(* Logix 5000 project; controller TFF vendor 1 type 14 code 107 rev 34.11; software revision 34.03; part 20 of 36 *)
(* tags used below, declared in another part *)
   Address : DINT;   // Temp Address
   Config : Configuration;   // Index Array used in configuration routines
   Index : DINT;   // Index
   NewSystem : DINT;
   AI101 : ALIAS FOR AnalogPoint[10];   // Filtrate Conductivity
   AI101_SIG : ALIAS FOR DigitalPoint[90];
   AI102 : ALIAS FOR AnalogPoint[11];   // Filtrate UV
   AI102_SIG : ALIAS FOR DigitalPoint[91];
   AI103 : ALIAS FOR AnalogPoint[12];   // Filtrate UV
   AI103_SIG : ALIAS FOR DigitalPoint[92];
   AI104 : ALIAS FOR AnalogPoint[9];   // Filtrate pH
   AI104_SIG : ALIAS FOR DigitalPoint[105];
   AlarmAnalog : AlarmAnalog[50];   // Analog Alarm Array
   AlarmControl : AlarmControl;   // Alarm Control
   AlarmDeviation : AlarmDeviation[20];   // Control Loop Deviation Alarm Array
   AnalogOutput : AnalogOutput[25];   // Analog Output Array
   AnalogPoint : AnalogInput[50];   // Analog Input Array
   Concentration : Concentration;
   ControlLoop : ControlLoop[20];   // Control Loop Array
   ControlLoop_FeedBagLevel : ALIAS FOR ControlLoop[2];   // Feed Bag Level Control Loop
   Diafiltration : Diafiltration;
   DigitalOutput : BOOL[256];   // Digital Output Array these bits are sent to output cards.
   DigitalPoint : DigitalPoint[150];   // Digital Point Array
   DP : ALIAS FOR AnalogPoint[40];   // Differential Pressure
   Drive : Drive[11];   // Drives Array
   ES001 : ALIAS FOR DigitalPoint[3];   // Emergency Stop
   FI001 : ALIAS FOR AnalogPoint[42];   // Feed Flow
   FI003 : ALIAS FOR AnalogPoint[17];
   FI003_SIG : ALIAS FOR DigitalPoint[106];
   FI003Alarm : ALIAS FOR AlarmAnalog[17];
   FI101 : ALIAS FOR AnalogPoint[2];   // Filtrate Flow
   FI101_SIG : ALIAS FOR DigitalPoint[93];
   FI101Alarm : ALIAS FOR AlarmAnalog[2];   // Filtrate Flow Alarm
   FI401 : ALIAS FOR AnalogPoint[43];   // Transfer Pump Flow
   LI001 : ALIAS FOR AnalogPoint[44];   // Feed Bag Volume
   LI001Alarm : ALIAS FOR AlarmAnalog[44];   // Feed Bag Volume Alarm
   MIX001 : ALIAS FOR AnalogPoint[14];   // Mixer Speed
   MIX001_SIG : ALIAS FOR DigitalPoint[104];
   Mixer : Mixer;   // Mixer config. structure
   NWP : ALIAS FOR AnalogPoint[45];   // Normalized Water Permeability
   Options : Options;   // Options List
   PCV001 : ALIAS FOR AnalogPoint[3];   // Retentate Pressure Control Valve Position
   PCV001_Control : PCV_Control;   // PCV001 Control UDT
   PCV001_SIG : ALIAS FOR DigitalPoint[102];
   PCV101 : ALIAS FOR AnalogPoint[4];   // Filtrate Pressure Control Valve Position
   PCV101_Control : PCV_Control;   // PCV101 Control UDT
   PCV101_SIG : ALIAS FOR DigitalPoint[103];
   PERM : ALIAS FOR AnalogPoint[46];   // Membrane Permeability
   PI001 : ALIAS FOR AnalogPoint[5];   // Feed Pressure
   PI001_SIG : ALIAS FOR DigitalPoint[97];
   PI002 : ALIAS FOR AnalogPoint[6];   // Retentate Pressure
   PI002_SIG : ALIAS FOR DigitalPoint[98];
   PI101 : ALIAS FOR AnalogPoint[7];   // Filtrate Pressure
   PI101_SIG : ALIAS FOR DigitalPoint[99];
   PI401 : ALIAS FOR AnalogPoint[8];   // Transfer Pump Pressure
   PI401_SIG : ALIAS FOR DigitalPoint[100];
   PSH001 : ALIAS FOR DigitalPoint[4];   // Feed Pump High Pressure
   PSH401 : ALIAS FOR DigitalPoint[5];   // Transfer Pump High Pressure
   PSL602 : ALIAS FOR DigitalPoint[0];   // Valves Air Defect
   PSL603 : ALIAS FOR DigitalPoint[10];   // Manifold Valves Air Defect
   SIC001 : ALIAS FOR Drive[1];   // Feed Pump
   SIC001DF : ALIAS FOR DigitalPoint[8];   // Feed Pump Defect
   SIC002 : ALIAS FOR Drive[2];   // Transfer Pump
   SIC002DF : ALIAS FOR DigitalPoint[9];   // Transfer Pump Defect
   SIC003 : ALIAS FOR Drive[3];   // Mixer
   SIC003DF : ALIAS FOR DigitalPoint[14];   // Mixer Defect
   SRL001 : ALIAS FOR DigitalPoint[15];   // Tank Skid Remote / Standalone
   Tank : TankManagement;   // Tank Management
   ThisSystem : SystemType;
   TI001 : ALIAS FOR AnalogPoint[13];   // Feed Bag Temperature
   TI001_SIG : ALIAS FOR DigitalPoint[101];
   TMP : ALIAS FOR AnalogPoint[41];   // Trans-membrane Pressure
   Totalizer : Totalizers[20];   // Totalizers Array
   UserCr1 : ALIAS FOR DigitalPoint[65];   // User Critical Alarm 1
   UserCr2 : ALIAS FOR DigitalPoint[67];   // User Critical Alarm 2
   UserNCr1 : ALIAS FOR DigitalPoint[64];   // User Non Critical Alarm 1
   UserNCr2 : ALIAS FOR DigitalPoint[66];   // User Non Critical Alarm 2
   Valve : Valve[100];   // Valve Array
   WI001 : ALIAS FOR AnalogPoint[15];   // Feed Bag Weight
   WI001_SIG : ALIAS FOR DigitalPoint[94];
   WI001Alarm : ALIAS FOR AlarmAnalog[15];   // Feed Bag Weight Alarm
   WI101 : ALIAS FOR AnalogPoint[0];   // Filtrate Weight
   WI101_SIG : ALIAS FOR DigitalPoint[95];
   WI101Alarm : ALIAS FOR AlarmAnalog[0];   // Filtrate Weight Alarm
   WI102 : ALIAS FOR AnalogPoint[1];   // Customer Filtrate Weight
   WI102_SIG : ALIAS FOR DigitalPoint[96];
   WI102Alarm : ALIAS FOR AlarmAnalog[1];   // Customer Filtrate Weight Alarm
   XC102_3DF : ALIAS FOR DigitalPoint[13];   // C8000 Defect
   XS001 : ALIAS FOR DigitalPoint[1];   // Door Closed
   XS002 : ALIAS FOR DigitalPoint[6];   // Clamshell Locking 1 Closed
   XS003 : ALIAS FOR DigitalPoint[7];   // Clamshell Locking 2 Closed
   XS006 : ALIAS FOR DigitalPoint[2];   // Door to Frame Locking Closed
   XS011 : ALIAS FOR DigitalPoint[11];   // Pump P001 Type
   XS012 : ALIAS FOR DigitalPoint[12];   // Pump P002 Type
   YA01 : ALIAS FOR DigitalPoint[50];   // PC to PLC communication failure
   YA02 : ALIAS FOR DigitalPoint[51];   // CCP Runtime communication failure
   YA03 : ALIAS FOR DigitalPoint[52];   // Historical Data collection failure
   YA04 : ALIAS FOR DigitalPoint[53];   // Hard Drive Overload
   YA05 : ALIAS FOR DigitalPoint[54];   // Database Overload
   YA06 : ALIAS FOR DigitalPoint[55];   // Node 0 communication failure - Smart
   YA07 : ALIAS FOR DigitalPoint[56];   // Node 0 internal defect - Smart
   YA08 : ALIAS FOR DigitalPoint[57];   // Node 1 communication failure - Clamshell
   YA09 : ALIAS FOR DigitalPoint[58];   // Node 1 internal defect - Clamshell
   YA10 : ALIAS FOR DigitalPoint[59];   // PLC Program Major Fault
   YA11 : ALIAS FOR DigitalPoint[60];   // Database Corrupted
   YA12 : ALIAS FOR DigitalPoint[61];   // Unauthorized accesses
   YA13 : ALIAS FOR DigitalPoint[62];   // Tank Size Mismatch
   YA14 : ALIAS FOR DigitalPoint[63];   // SQL Server Write Failure
   YA15 : ALIAS FOR DigitalPoint[69];   // Node 3 Communication Failure - Pump
   YA16 : ALIAS FOR DigitalPoint[70];   // Node 3 Internal Defect - Pump
   YA17 : ALIAS FOR DigitalPoint[71];   // Node 4 Communication Failure - Instrum
   YA18 : ALIAS FOR DigitalPoint[72];   // Node 4 Internal Defect - Instrum
   YA19 : ALIAS FOR DigitalPoint[73];   // Node 5 Communication Failure - Tank
   YA20 : ALIAS FOR DigitalPoint[74];   // Node 5 Internal Defect - Tank
   YA21 : ALIAS FOR DigitalPoint[75];   // Node 6 IND331 Communication Failure
   YA22 : ALIAS FOR DigitalPoint[76];   // Node 7 IND131 Communication Failure
   YA41 : ALIAS FOR DigitalPoint[77];   // YA41 Operating Time Exceeded
   ZSDF : ALIAS FOR DigitalPoint[68];   // ZSDF Clamshell Locking Defect
(* Process, continued *)

ROUTINE Alarm_Init_Config   (* structured text *)
   (* =======================================================================
   	Alarm_Init_SP : initialized  parameter to default values
   
   	List of treatments
   		- Analog alarms set point with scale Min and Max
   		- Deviation alarms
   		- Digital alarmss
   		- Valves alarms
   	-----------------------------------------------------------------------------------------------------------------------------------------------------
   	History
   		2020-Sep-28 - Merck - Q.Spindler - Initial version for Candidate Release 3.00.00.01.a
   		2021-May-31 - DAVIDSON- Ch. ARBOGAST - Modifications for Candidate Release 3.01.00.00.a
   		On Analog Set point, add lines for set WI001 & LI001, HI & HIHI values according to actual tank size
   		On Analog Set point, add lines for set WI101 & WI102 & FI003 & FI101, HI & HIHI values according to actual system type
   		On Discrete Alarms: modify YA03.DelayTimerSP := 80
   		On Discrete Alarms: for all “_SIG” alarms, modify: Priority := 0 , DelayTimerSP := 10
   		On Discrete Alarms add line with WI001_SIG settings
   		On Discrete Alarms, last line FI003 settings: replace AI104 by FI003 (2x)
   =============================================================================================================================*)
   
   (*Analog Set point to min/max scale, Enable alarm, timer to  2s
   ============================================================*)
   	FOR Index := 0 to 49 by 1 do
   		IF AnalogPoint[Index].EnableCfg THEN
   			AlarmAnalog[Index].Override := 0; // Enable
   			AlarmAnalog[Index].LOLO := AnalogPoint[Index].ScaledMin ;
   			AlarmAnalog[Index].LO := AnalogPoint[Index].ScaledMin ;
   			AlarmAnalog[Index].HI := AnalogPoint[Index].ScaledMax ;
   			AlarmAnalog[Index].HIHI := AnalogPoint[Index].ScaledMax ;
   			AlarmAnalog[Index].LOLOTimerSP := 2 ;
   			AlarmAnalog[Index].LOTimerSP := 2 ;
   			AlarmAnalog[Index].HITimerSP := 2 ;
   			AlarmAnalog[Index].HIHITimerSP := 2 ;
   		END_IF;
   	End_for ;
   	(* Tank 60(50L) *)
   	IF Tank.Config.TankSelected = 1 THEN
   		WI001Alarm.HIHI := 60 ;
   		WI001Alarm.HI := 60 ;
   		LI001Alarm.HIHI := 50 ;
   		LI001Alarm.HI := 50 ;
   	END_IF ;
   	(* Tank 120(100L) *)
   	IF Tank.Config.TankSelected = 2 THEN
   		WI001Alarm.HIHI := 120 ;
   		WI001Alarm.HI := 120 ;
   		LI001Alarm.HIHI := 100 ;
   		LI001Alarm.HI := 100 ;
   	END_IF ;
   	(* Tank 240(200L) *)
   	IF Tank.Config.TankSelected = 3 THEN
   		WI001Alarm.HIHI := 240 ;
   		WI001Alarm.HI := 240 ;
   		LI001Alarm.HIHI := 200 ;
   		LI001Alarm.HI := 200 ;
   	END_IF ;
   	(* TF2S *)
   	IF NewSystem = 123 THEN
   		WI101Alarm.HIHI := 600 ;
   		WI101Alarm.HI := 600 ;
   		WI102Alarm.HIHI := 1000 ;
   		WI102Alarm.HI := 1000 ;
   		FI003Alarm.HIHI := 15 ;
   		FI003Alarm.HI := 15 ;
   		FI101Alarm.HIHI := 15 ;
   		FI101Alarm.HI := 15 ;
   	END_IF ;
   	(* TF3S *)
   	IF NewSystem = 124 THEN
   		WI101Alarm.HIHI := 1500 ;
   		WI101Alarm.HI := 1500 ;
   		WI102Alarm.HIHI := 1500 ;
   		WI102Alarm.HI := 1500 ;
   		FI003Alarm.HIHI := 25 ;
   		FI003Alarm.HI := 25 ;
   		FI101Alarm.HIHI := 25 ;
   		FI101Alarm.HI := 25 ;
   	END_IF ;
   
   (*Deviation alarm HI 100% HIHI 100%, Disable alarm, timer to 2s
   ============================================================*)
   	FOR Index := 0 to 19 by 1 do
   		IF AlarmDeviation[Index].EnableCfg THEN
   			AlarmDeviation[Index].Override := 1; // Disable
   			AlarmDeviation[Index].HI := 100 ;
   			AlarmDeviation[Index].HIHI := 100 ;
   			AlarmDeviation[Index].HITimerSP := 2 ;
   			AlarmDeviation[Index].HIHITImerSP := 2 ;
   		END_IF;
   	End_for ;
   
   (* Discrete Alarms
   ============================================================*)
   	ES001.DelayTimerSP := 0;
   	PSH001.Override := 0; PSH001.Priority := 1; PSH001.DelayTimerSP := 0;
   	PSH401.Override := 0; PSH401.Priority := 1; PSH401.DelayTimerSP := 0;
   	PSL602.Override := 0; PSL602.Priority := 1; PSL602.DelayTimerSP := 2;
   	SIC001DF.Override := 0; SIC001DF.Priority := 1; SIC001DF.DelayTimerSP :=1;
   	SIC002DF.Override := 0; SIC002DF.Priority := 1; SIC002DF.DelayTimerSP :=1;
   	SIC003DF.Override := 0; SIC003DF.Priority := 1; SIC003DF.DelayTimerSP :=1;
   	XC102_3DF.Override := 0; XC102_3DF.Priority := 1; XC102_3DF.DelayTimerSP :=1;
   	ZSDF.Override := 0; ZSDF.Priority := 1; ZSDF.DelayTimerSP :=1;
   	XS001.Override := 0; XS001.Priority := 1; XS001.DelayTimerSP :=1;
   	PSL603.Override := 0; PSL603.Priority := 1; PSL603.DelayTimerSP :=1;
   
   	YA01.Override := 0; YA01.Priority := 0; YA01.DelayTimerSP := 60;
   	YA02.Override := 0; YA02.Priority := 0; YA02.DelayTimerSP := 60;
   	YA03.Override := 0; YA03.Priority := 0; YA03.DelayTimerSP := 80;
   	YA04.Override := 0; YA04.Priority := 0; YA04.DelayTimerSP := 60;
   	YA05.Override := 0; YA05.Priority := 0; YA05.DelayTimerSP := 60;
   	YA06.Override := 0; YA06.Priority := 1; YA06.DelayTimerSP := 5;
   	YA07.Override := 0; YA07.Priority := 0; YA07.DelayTimerSP := 2;
   	YA08.Override := 0; YA08.Priority := 1; YA08.DelayTimerSP := 5;
   	YA09.Override := 0; YA09.Priority := 0; YA09.DelayTimerSP := 2;
   	YA10.DelayTimerSP := 0;
   	YA11.Override := 1; YA11.Priority := 0; YA11.DelayTimerSP := 5;
   	YA12.Override := 0; YA12.Priority := 0; YA12.DelayTimerSP := 0;
   	YA13.Override := 0; YA13.Priority := 0; YA13.DelayTimerSP := 2;
   	YA14.Override := 0; YA14.Priority := 0; YA14.DelayTimerSP := 60;
   	YA15.Override := 0; YA15.Priority := 1; YA15.DelayTimerSP := 5;
   	YA16.Override := 0; YA16.Priority := 0; YA16.DelayTimerSP := 2;
   	YA17.Override := 0; YA17.Priority := 1; YA17.DelayTimerSP := 5;
   	YA18.Override := 0; YA18.Priority := 0; YA18.DelayTimerSP := 2;
   	YA19.Override := 0; YA19.Priority := 1; YA19.DelayTimerSP := 5;
   	YA20.Override := 0; YA20.Priority := 0; YA20.DelayTimerSP := 2;
   	YA21.Override := 0; YA21.Priority := 1; YA21.DelayTimerSP := 5;
   	YA22.Override := 0; YA22.Priority := 1; YA22.DelayTimerSP := 5;
   
   	AI101_SIG.Override := 0; AI101_SIG.Priority := 0; AI101_SIG.DelayTimerSP := 10;
   	AI102_SIG.Override := 0; AI102_SIG.Priority := 0; AI102_SIG.DelayTimerSP := 10;
   	AI103_SIG.Override := 0; AI103_SIG.Priority := 0; AI103_SIG.DelayTimerSP := 10;
   	FI101_SIG.Override := 0; FI101_SIG.Priority := 0; FI101_SIG.DelayTimerSP := 10;
   	WI001_SIG.Override := 0; WI001_SIG.Priority := 0; WI001_SIG.DelayTimerSP := 10;
   	WI101_SIG.Override := 0; WI101_SIG.Priority := 0; WI101_SIG.DelayTimerSP := 10;
   	WI102_SIG.Override := 0; WI102_SIG.Priority := 0; WI102_SIG.DelayTimerSP := 10;
   	PI001_SIG.Override := 0; PI001_SIG.Priority := 0; PI001_SIG.DelayTimerSP := 10;
   	PI002_SIG.Override := 0; PI002_SIG.Priority := 0; PI002_SIG.DelayTimerSP := 10;
   	PI101_SIG.Override := 0; PI101_SIG.Priority := 0; PI101_SIG.DelayTimerSP := 10;
   	PI401_SIG.Override := 0; PI401_SIG.Priority := 0; PI401_SIG.DelayTimerSP := 10;
   	TI001_SIG.Override := 0; TI001_SIG.Priority := 0; TI001_SIG.DelayTimerSP := 10;
   	PCV001_SIG.Override := 0; PCV001_SIG.Priority := 0; PCV001_SIG.DelayTimerSP := 10;
   	PCV101_SIG.Override := 0; PCV101_SIG.Priority := 0; PCV101_SIG.DelayTimerSP := 10;
   	MIX001_SIG.Override := 0; MIX001_SIG.Priority := 0; MIX001_SIG.DelayTimerSP := 10;
   	AI104_SIG.Override := 0; AI104_SIG.Priority := 0; AI104_SIG.DelayTimerSP := 10;
   	FI003_SIG.Override := 0; FI003_SIG.Priority := 0; FI003_SIG.DelayTimerSP := 10;
   
   	UserNCr1.Priority := 0; UserNCr1.DelayTimerSP := 0;
   	UserCr1.Priority := 1; UserCr1.DelayTimerSP := 0;
   	UserNCr2.Priority := 0; UserNCr2.DelayTimerSP := 0;
   	UserCr2.Priority := 1; UserCr2.DelayTimerSP := 0;
   
   // Reset Init command
   AlarmControl.InitAlarmConfig := 0;
END_ROUTINE

ROUTINE Concentration_Diafiltration   (* ladder *)
// Agitator Control Routine
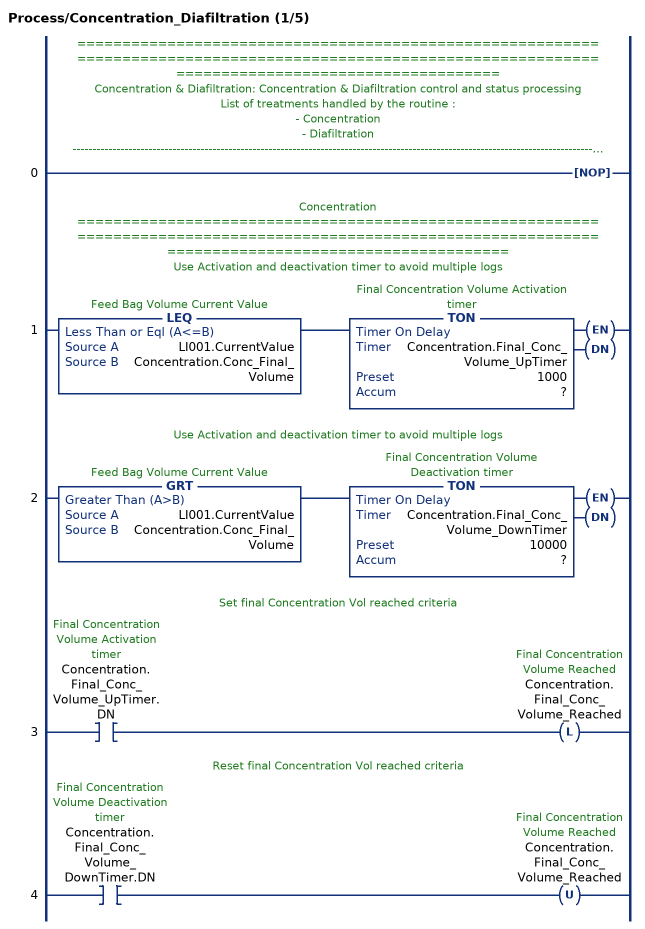
   // ========================================================================================================================================================
   //                                                                                                    Concentration & Diafiltration: Concentration & Diafiltration control and status processing
   //                                                     List of treatments handled by the routine :
   //                                                          - Concentration
   //                                                          - Diafiltration
   //                                                     -----------------------------------------------------------------------------------------------------------------------------------------------------
   //                                                     History
   //                                                          2019-AUG-13 - Actemium - B. Roch - Initial version for Candidate Release 3.00.00.00.a
   //                                                           2020-SEP-24 - Merck - Q. Spindler - Modifications for Candidate Release 3.00.00.01.a
   //                                        - Add Timer for activation and deactivation of Volume/Protein reached status to avoid unwanted logs
   // ========================================================================================================================================================
   0: NOP();
   // Concentration
   // ==========================================================================================================================================================
   // Use Activation and deactivation timer to avoid multiple logs
   1: LEQ(LI001.CurrentValue,Concentration.Conc_Final_Volume)TON(Concentration.Final_Conc_Volume_UpTimer,?,?);
   // Use Activation and deactivation timer to avoid multiple logs
   2: GRT(LI001.CurrentValue,Concentration.Conc_Final_Volume)TON(Concentration.Final_Conc_Volume_DownTimer,?,?);
   // Set final Concentration Vol reached criteria
   3: XIC(Concentration.Final_Conc_Volume_UpTimer.DN)OTL(Concentration.Final_Conc_Volume_Reached);
   // Reset final Concentration Vol reached criteria
   4: XIC(Concentration.Final_Conc_Volume_DownTimer.DN)OTU(Concentration.Final_Conc_Volume_Reached);
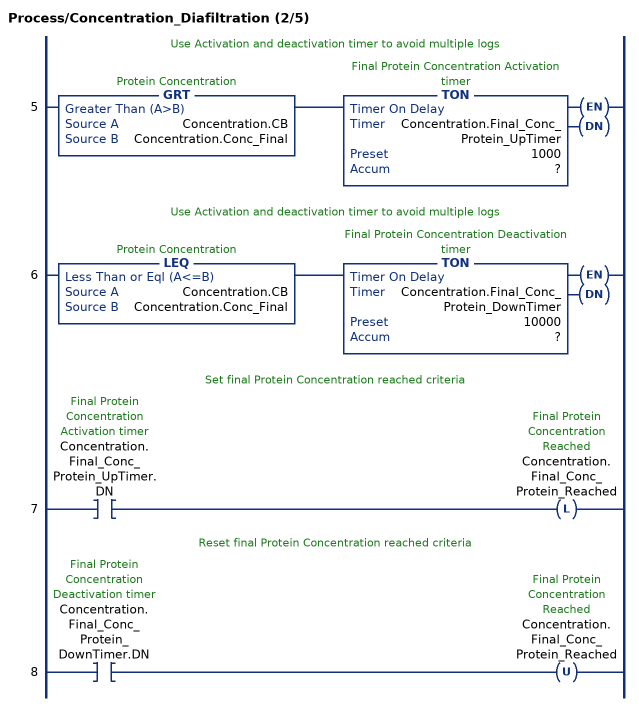
   // Use Activation and deactivation timer to avoid multiple logs
   5: GRT(Concentration.CB,Concentration.Conc_Final)TON(Concentration.Final_Conc_Protein_UpTimer,?,?);
   // Use Activation and deactivation timer to avoid multiple logs
   6: LEQ(Concentration.CB,Concentration.Conc_Final)TON(Concentration.Final_Conc_Protein_DownTimer,?,?);
   // Set final Protein Concentration reached criteria
   7: XIC(Concentration.Final_Conc_Protein_UpTimer.DN)OTL(Concentration.Final_Conc_Protein_Reached);
   // Reset final Protein Concentration reached criteria
   8: XIC(Concentration.Final_Conc_Protein_DownTimer.DN)OTU(Concentration.Final_Conc_Protein_Reached);
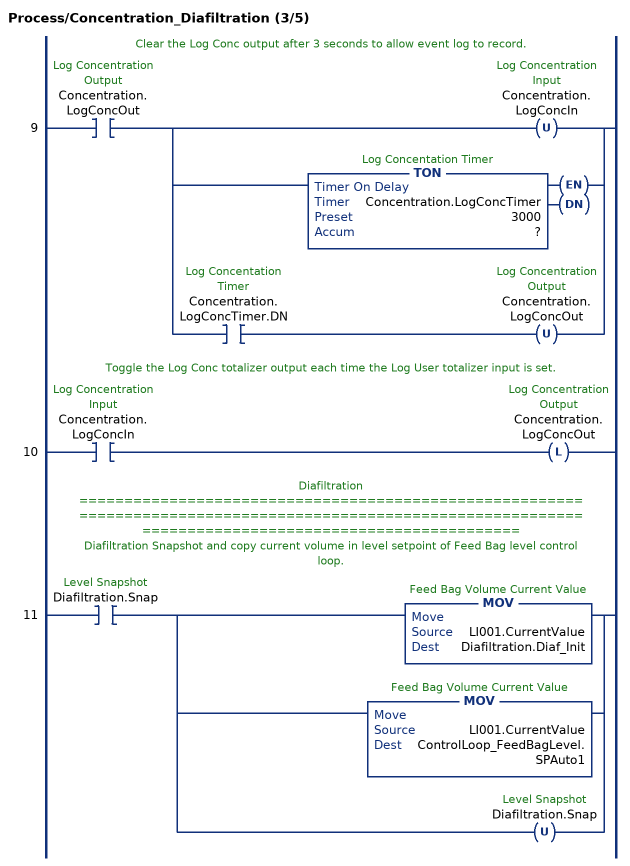
   // Clear the Log Conc output after 3 seconds to allow event log to record.
   9: XIC(Concentration.LogConcOut)[OTU(Concentration.LogConcIn) ,TON(Concentration.LogConcTimer,?,?) ,XIC(Concentration.LogConcTimer.DN) OTU(Concentration.LogConcOut) ];
   // Toggle the Log Conc totalizer output each time the Log User totalizer input is set.
   10: XIC(Concentration.LogConcIn)OTL(Concentration.LogConcOut);
   // Diafiltration
   // ==========================================================================================================================================================
   // Diafiltration Snapshot and copy current volume in level setpoint of Feed Bag level control loop.
   11: XIC(Diafiltration.Snap)[MOV(LI001.CurrentValue,Diafiltration.Diaf_Init) ,MOV(LI001.CurrentValue,ControlLoop_FeedBagLevel.SPAuto1) ,OTU(Diafiltration.Snap) ];
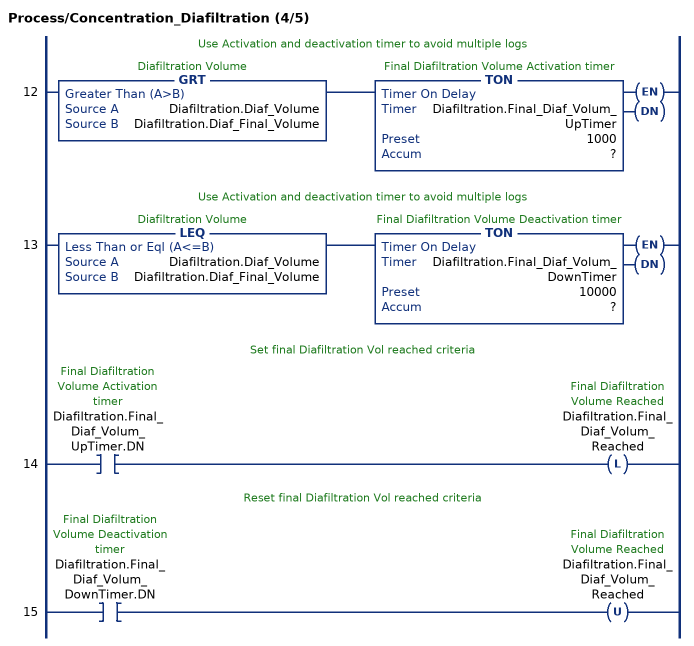
   // Use Activation and deactivation timer to avoid multiple logs
   12: GRT(Diafiltration.Diaf_Volume,Diafiltration.Diaf_Final_Volume)TON(Diafiltration.Final_Diaf_Volum_UpTimer,?,?);
   // Use Activation and deactivation timer to avoid multiple logs
   13: LEQ(Diafiltration.Diaf_Volume,Diafiltration.Diaf_Final_Volume)TON(Diafiltration.Final_Diaf_Volum_DownTimer,?,?);
   // Set final Diafiltration Vol reached criteria
   14: XIC(Diafiltration.Final_Diaf_Volum_UpTimer.DN)OTL(Diafiltration.Final_Diaf_Volum_Reached);
   // Reset final Diafiltration Vol reached criteria
   15: XIC(Diafiltration.Final_Diaf_Volum_DownTimer.DN)OTU(Diafiltration.Final_Diaf_Volum_Reached);
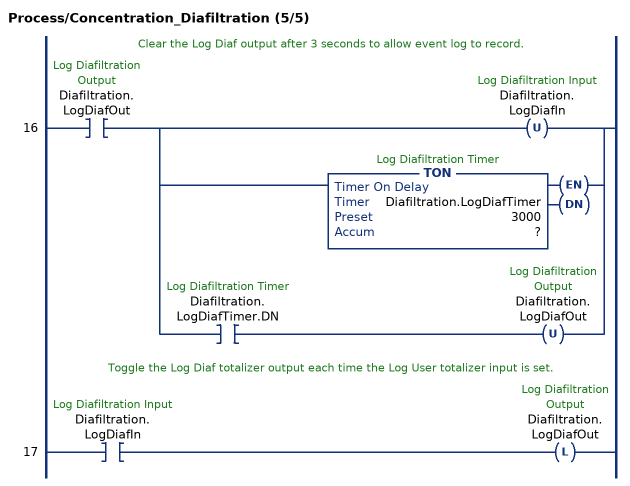
   // Clear the Log Diaf output after 3 seconds to allow event log to record.
   16: XIC(Diafiltration.LogDiafOut)[OTU(Diafiltration.LogDiafIn) ,TON(Diafiltration.LogDiafTimer,?,?) ,XIC(Diafiltration.LogDiafTimer.DN) OTU(Diafiltration.LogDiafOut) ];
   // Toggle the Log Diaf totalizer output each time the Log User totalizer input is set.
   17: XIC(Diafiltration.LogDiafIn)OTL(Diafiltration.LogDiafOut);
END_ROUTINE

ROUTINE Config_AnalogOutput   (* structured text *)
   (* ==========================================================
   	Config AnalogOutput : Configure AnalogOutput Structure
   
   	List of treatments
   		- AnalogOutput[0] : Retentate Pressure Control Valve Setpoint
   		- AnalogOutput[1] : Filtrate Pressure Control Valve Setpoint
   		- AnalogOutput[2] : Feed Pump Speed Setpoint
   		- AnalogOutput[3] : Transfer Pump Speed Setpoint
   		- AnalogOutput[4] : Mixer Speed Setpoint
   		- Reset Loop : Set to 0 the AnalogOutput[5 to 24].EnableCfg
   
   -----------------------------------------------------------------------------------------------------------------------------------------------------
   	History
   		2019-AUG-13 - ACTEMIUM - B. Roch - Initial version for Candidate Release 3.00.00.00.a
   ============================================================*)
   
   (*AnalogOutput[0] : PCV001 Retentate Pressure Control Valve Setpoint
   ============================================================*)
   AnalogOutput[0].EnableCfg := 1 ;
   AnalogOutput[0].RawMin := 0 ;
   AnalogOutput[0].RawMax := 2047 ;
   AnalogOutput[0].ScaledMin := 0 ;
   AnalogOutput[0].ScaledMax := 100 ;
   
   (*AnalogOutput[1] : PCV101 Filtrate Pressure Control Valve Setpoint
   ============================================================*)
   AnalogOutput[1].EnableCfg := 1 ;
   AnalogOutput[1].RawMin := 0 ;
   AnalogOutput[1].RawMax := 2047 ;
   AnalogOutput[1].ScaledMin := 0 ;
   AnalogOutput[1].ScaledMax := 100 ;
   
   (*AnalogOutput[2] : SIC001 Feed Pump Speed Setpoint
   ============================================================*)
   AnalogOutput[2].EnableCfg := 1 ;
   AnalogOutput[2].RawMin := 0 ;
   AnalogOutput[2].RawMax := 27648 ;
   AnalogOutput[2].ScaledMin := 0 ;
   AnalogOutput[2].ScaledMax := 100 ;
   
   (*AnalogOutput[3] : SIC002 Transfer Pump Speed Setpoint
   ============================================================*)
   AnalogOutput[3].EnableCfg := 1 ;
   AnalogOutput[3].RawMin := 0 ;
   AnalogOutput[3].RawMax := 27648 ;
   AnalogOutput[3].ScaledMin := 0 ;
   AnalogOutput[3].ScaledMax := 100 ;
   
   (*AnalogOutput[4] : SIC003 Mixer Speed Setpoint
   ============================================================*)
   AnalogOutput[4].EnableCfg := 1 ;
   AnalogOutput[4].RawMin := 0 ;
   AnalogOutput[4].RawMax := 2047 ;
   AnalogOutput[4].ScaledMin := 0 ;
   AnalogOutput[4].ScaledMax := 100 ;
   
   
   (*Reset Loop : Set to 0 the AnalogOutput[12 to 24].EnableCfg
   ============================================================*)
   FOR Config.IndexA0 := 5 to 24 by 1 do
   	AnalogOutput[Config.IndexA0].EnableCfg := 0 ;
   End_for ;
   
END_ROUTINE

ROUTINE Config_AnalogPoint   (* structured text *)
// Apply the default configuration
   (* ==========================================================
   	Config AnalogPoint : Configure AnalogPoint Structure
   
   	List of treatments
   		- AnalogPoint[0] : Filtrate Weight WI101
   		- AnalogPoint[1] : Customer Filtrate Weight WI102
   		- AnalogPoint[2] : Filtrate Flow FI101
   		- AnalogPoint[3] : Retentate Pressure Control Valve Position PCV001
   		- AnalogPoint[4] : Filtrate Pressure Control Valve Position PCV101
   		- AnalogPoint[5] : Feed Pressure PI001
   		- AnalogPoint[6] : Retentate Pressure PI002
   		- AnalogPoint[7] : Filtrate Pressure PI101
   		- AnalogPoint[8] : Transfer Pump Pressure PI401
   		- AnalogPoint[9] : Filtrate pH AI104
   		- AnalogPoint[10]: Filtrate Conductivity AI101
   		- AnalogPoint[11]: Filtrate UV AI102
   		- AnalogPoint[12]: Filtrate UV AI103
   		- AnalogPoint[13]: Feed Bag Temperature TI001
   		- AnalogPoint[14]: Mixer Speed MIX001
   		- AnalogPoint[15]: Feed Bag Weight WI001
   		- AnalogPoint[16]: Spare
   		- AnalogPoint[17]: Retentate Flow FI003
   		- Reset Loop : Set to 0 the AnalogPoint[18 to 39].EnableCfg
   		- AnalogPoint[40]: Differential Pressure DP
   		- AnalogPoint[41]: Trans-Membrane Pressure TMP
   		- AnalogPoint[42]: Feed Flow FI001
   		- AnalogPoint[43]: Transfer Pump Flow FI401
   		- AnalogPoint[44]: Feed Bag Volume LI001
   		- AnalogPoint[45]: Normalized Water Permeability NWP
   		- AnalogPoint[46]: Membrane Permeability PERM
   		- Reset Loop : Set to 0 the AnalogPoint[47 to 49].EnableCfg
   
   -----------------------------------------------------------------------------------------------------------------------------------------------------
   	History
   		2019-AUG-13 - ACTEMIUM - B. Roch - Initial version for Candidate Release 3.00.00.00.a
   		2019-SEP-26 - ACTEMIUM - B. Roch - Modifications for Candidate Release 3.00.00.00.c
   					- Change RealCfg to 1 for AI101
   					- delete the enableCfg for AI101 outside the option check
   		2020-SEP-29 - Merck - Q. Spindler - Modifications for Candidate Release 3.00.00.01.a
   					- Add FI003
   		2020-NOV-24 - Merck - Q. Spindler - Modifications for Candidate Release 3.00.00.01.b
   					- Change FI003 option
   ============================================================*)
   
   
   (*AnalogPoint[0] : Filtrate Weight WI101
   ============================================================*)
   
   IF Options.No_Filtrate_Measurement OR Options.WI102 OR Options.FI101 OR Options.WI102_FI101 THEN
   	AnalogPoint[0].EnableCfg := 0 ;
   	AlarmAnalog[0].EnableCfg := 0 ;
   ELSIF Options.WI101 OR Options.WI101_FI101 THEN
   	AnalogPoint[0].EnableCfg := 1 ;
   	AlarmAnalog[0].EnableCfg := 1 ;
   ELSE
   	AnalogPoint[0].EnableCfg := 0 ;
   	AlarmAnalog[0].EnableCfg := 0 ;
   END_IF;
   
   AnalogPoint[0].Address := 0 ;
   AnalogPoint[0].RealCfg := 0 ;
   AnalogPoint[0].RawMin := 0 ;
   AnalogPoint[0].RawMax := 99999 ;
   AnalogPoint[0].OverrideCfg := 1 ;
   AnalogPoint[0].ScaledMin := 0;
   AnalogPoint[0].ScaledMax := 9999.9;
   AlarmAnalog[0].FeedPumpEnable := 0 ;
   AlarmAnalog[0].FeedPumpTag := 0 ;
   AlarmAnalog[0].TransferPumpEnable := 0 ;
   AlarmAnalog[0].TransferPumpTag := 0 ;
   AlarmAnalog[0].Disable := 0 ;
   AlarmAnalog[0].HIHIEnable := 0 ;
   
   
   (*AnalogPoint[1] : Customer Filtrate Weight WI102
   ============================================================*)
   
   IF Options.No_Filtrate_Measurement OR Options.WI101 OR Options.FI101 OR Options.WI101_FI101 THEN
   	AnalogPoint[1].EnableCfg := 0 ;
   	AlarmAnalog[1].EnableCfg := 0 ;
   ELSIF Options.WI102 OR Options.WI102_FI101 THEN
   	AnalogPoint[1].EnableCfg := 1 ;
   	AlarmAnalog[1].EnableCfg := 1 ;
   ELSE
   	AnalogPoint[1].EnableCfg := 0 ;
   	AlarmAnalog[1].EnableCfg := 0 ;
   END_IF;
   
   AnalogPoint[1].Address := 1 ;
   AnalogPoint[1].RawMin := 6553 ;
   AnalogPoint[1].RawMax := 32767 ;
   AnalogPoint[1].RealCfg := 0 ;
   AnalogPoint[1].OverrideCfg := 1 ;
   AlarmAnalog[1].FeedPumpEnable := 0 ;
   AlarmAnalog[1].FeedPumpTag := 0 ;
   AlarmAnalog[1].TransferPumpEnable := 0 ;
   AlarmAnalog[1].TransferPumpTag := 0 ;
   AlarmAnalog[1].Disable := 0 ;
   AlarmAnalog[1].HIHIEnable := 0 ;
   
   (*AnalogPoint[2] : Filtrate Flow FI101 (Flow Meter)
   ============================================================*)
   
   IF Options.No_Filtrate_Measurement THEN
   	AnalogPoint[2].EnableCfg := 0 ;
   	AlarmAnalog[2].EnableCfg := 0 ;
   	AnalogPoint[2].RealCfg := 1 ;
   ELSIF Options.WI102 OR Options.WI101 THEN
   	AnalogPoint[2].EnableCfg := 1 ;
   	AlarmAnalog[2].EnableCfg := 1 ;
   	AnalogPoint[2].RealCfg := 0 ;
   ELSIF Options.FI101 OR Options.WI101_FI101 OR Options.WI102_FI101 THEN
   	AnalogPoint[2].EnableCfg := 1 ;
   	AlarmAnalog[2].EnableCfg := 1 ;
   	AnalogPoint[2].RealCfg := 1 ;
   ELSE
   	AnalogPoint[2].EnableCfg := 0 ;
   	AlarmAnalog[2].EnableCfg := 0 ;
   	AnalogPoint[2].RealCfg := 1 ;
   END_IF;
   
   AnalogPoint[2].Address := 2 ;
   AnalogPoint[2].RawMin := 6553 ;
   AnalogPoint[2].RawMax := 32767 ;
   AnalogPoint[2].OverrideCfg := 1 ;
   AlarmAnalog[2].FeedPumpEnable := 1 ;
   AlarmAnalog[2].FeedPumpTag := 1 ;
   AlarmAnalog[2].TransferPumpEnable := 0 ;
   AlarmAnalog[2].TransferPumpTag := 0 ;
   AlarmAnalog[2].Disable := 0 ;
   AlarmAnalog[2].HIHIEnable := 0 ;
   
   (*AnalogPoint[3] : Retentate Pressure Control Valve Position PCV001
   ============================================================*)
   AnalogPoint[3].EnableCfg := 1 ;
   AnalogPoint[3].Address := 3 ;
   AnalogPoint[3].RawMin := 6553 ;
   AnalogPoint[3].RawMax := 32767 ;
   AnalogPoint[3].RealCfg := 0 ;
   AnalogPoint[3].OverrideCfg := 0 ;
   AlarmAnalog[3].FeedPumpEnable := 0 ;
   AlarmAnalog[3].FeedPumpTag := 0 ;
   AlarmAnalog[3].TransferPumpEnable := 0 ;
   AlarmAnalog[3].TransferPumpTag := 0 ;
   AlarmAnalog[3].EnableCfg := 0 ;
   AlarmAnalog[3].Disable := 0 ;
   AlarmAnalog[3].HIHIEnable := 0 ;
   
   (*AnalogPoint[4] : Filtrate Pressure Control Valve Position PCV101
   ============================================================*)
   AnalogPoint[4].EnableCfg := 1 ;
   AnalogPoint[4].Address := 4 ;
   AnalogPoint[4].RawMin := 6553 ;
   AnalogPoint[4].RawMax := 32767 ;
   AnalogPoint[4].RealCfg := 0 ;
   AnalogPoint[4].OverrideCfg := 0 ;
   AlarmAnalog[4].FeedPumpEnable := 0 ;
   AlarmAnalog[4].FeedPumpTag := 0 ;
   AlarmAnalog[4].TransferPumpEnable := 0 ;
   AlarmAnalog[4].TransferPumpTag := 0 ;
   AlarmAnalog[4].EnableCfg := 0 ;
   AlarmAnalog[4].Disable := 0 ;
   AlarmAnalog[4].HIHIEnable := 0 ;
   
   (*AnalogPoint[5] : Feed Pressure PI001
   ============================================================*)
   AnalogPoint[5].EnableCfg := 1 ;
   AnalogPoint[5].Address := 5 ;
   AnalogPoint[5].RawMin := 6553 ;
   AnalogPoint[5].RawMax := 32767 ;
   AnalogPoint[5].RealCfg := 1 ;
   AnalogPoint[5].OverrideCfg := 1 ;
   AlarmAnalog[5].FeedPumpEnable := 1 ;
   AlarmAnalog[5].FeedPumpTag := 1 ;
   AlarmAnalog[5].TransferPumpEnable := 0 ;
   AlarmAnalog[5].TransferPumpTag := 0 ;
   AlarmAnalog[5].EnableCfg := 1 ;
   AlarmAnalog[5].Disable := 0 ;
   AlarmAnalog[5].HIHIEnable := 1 ;
   
   (*AnalogPoint[6] : Retentate Pressure PI002
   ============================================================*)
   AnalogPoint[6].EnableCfg := 1 ;
   AlarmAnalog[6].EnableCfg := 1 ;
   AnalogPoint[6].Address := 6 ;
   AnalogPoint[6].RawMin := 6553 ;
   AnalogPoint[6].RawMax := 32767 ;
   AnalogPoint[6].RealCfg := 1 ;
   AnalogPoint[6].OverrideCfg := 1 ;
   AlarmAnalog[6].FeedPumpEnable := 1 ;
   AlarmAnalog[6].FeedPumpTag := 1 ;
   AlarmAnalog[6].TransferPumpEnable := 0 ;
   AlarmAnalog[6].TransferPumpTag := 0 ;
   AlarmAnalog[6].Disable := 0 ;
   AlarmAnalog[6].HIHIEnable := 1 ;
   
   (*AnalogPoint[7] : Filtrate Pressure PI101
   ============================================================*)
   AnalogPoint[7].EnableCfg := 1 ;
   AlarmAnalog[7].EnableCfg := 1 ;
   AnalogPoint[7].Address := 7 ;
   AnalogPoint[7].RawMin := 6553 ;
   AnalogPoint[7].RawMax := 32767 ;
   AnalogPoint[7].RealCfg := 1 ;
   AnalogPoint[7].OverrideCfg := 1 ;
   AlarmAnalog[7].FeedPumpEnable := 1 ;
   AlarmAnalog[7].FeedPumpTag := 1 ;
   AlarmAnalog[7].TransferPumpEnable := 0 ;
   AlarmAnalog[7].TransferPumpTag := 0 ;
   AlarmAnalog[7].Disable := 0 ;
   AlarmAnalog[7].HIHIEnable := 1 ;
   
   (*AnalogPoint[8] : Transfer Pump Pressure PI401
   ============================================================*)
   AnalogPoint[8].EnableCfg := 1 ;
   AlarmAnalog[8].EnableCfg := 1 ;
   AnalogPoint[8].Address := 8 ;
   AnalogPoint[8].RawMin := 6553 ;
   AnalogPoint[8].RawMax := 32767 ;
   AnalogPoint[8].RealCfg := 1 ;
   AnalogPoint[8].OverrideCfg := 1 ;
   AlarmAnalog[8].FeedPumpEnable := 0 ;
   AlarmAnalog[8].FeedPumpTag := 0 ;
   AlarmAnalog[8].TransferPumpEnable := 1 ;
   AlarmAnalog[8].TransferPumpTag := 2 ;
   AlarmAnalog[8].Disable := 0 ;
   AlarmAnalog[8].HIHIEnable := 1 ;
   
   (*AnalogPoint[9] : Filtrate pH AI104
   ============================================================*)
   
   IF Options.No_Device_Connected OR Options.AI102_AI103 OR Options.AI101 OR Options.AI101_AI102_AI103 THEN
   	AnalogPoint[9].EnableCfg := 0 ;
   	AlarmAnalog[9].EnableCfg := 0 ;
   ELSIF Options.AI101_AI104 OR Options.AI101_AI102_AI103_AI104 THEN
   	AnalogPoint[9].EnableCfg := 1 ;
   	AlarmAnalog[9].EnableCfg := 1 ;
   ELSE
   	AnalogPoint[9].EnableCfg := 0 ;
   	AlarmAnalog[9].EnableCfg := 0 ;
   END_IF;
   
   AnalogPoint[9].Address := 9 ;
   AnalogPoint[9].RawMin := 6553 ;
   AnalogPoint[9].RawMax := 32767 ;
   AnalogPoint[9].RealCfg := 1 ;
   AnalogPoint[9].OverrideCfg := 1 ;
   AlarmAnalog[9].FeedPumpEnable := 0 ;
   AlarmAnalog[9].FeedPumpTag := 0 ;
   AlarmAnalog[9].TransferPumpEnable := 0 ;
   AlarmAnalog[9].TransferPumpTag := 0 ;
   AlarmAnalog[9].Disable := 0 ;
   AlarmAnalog[9].HIHIEnable := 0 ;
   
   (*AnalogPoint[10]: Filtrate Conductivity AI101
   ============================================================*)
   
   IF Options.No_Device_Connected OR Options.AI102_AI103 THEN
   	AnalogPoint[10].EnableCfg := 0 ;
   	AlarmAnalog[10].EnableCfg := 0 ;
   ELSIF Options.AI101 OR Options.AI101_AI102_AI103  OR Options.AI101_AI104 OR Options.AI101_AI102_AI103_AI104 THEN
   	AnalogPoint[10].EnableCfg := 1 ;
   	AlarmAnalog[10].EnableCfg := 1 ;
   ELSE
   	AnalogPoint[10].EnableCfg := 0 ;
   	AlarmAnalog[10].EnableCfg := 0 ;
   END_IF;
   
   AnalogPoint[10].Address := 10 ;
   AnalogPoint[10].RawMin := 6553 ;
   AnalogPoint[10].RawMax := 32767 ;
   AnalogPoint[10].RealCfg := 1 ;
   AnalogPoint[10].OverrideCfg := 1 ;
   AlarmAnalog[10].FeedPumpEnable := 0 ;
   AlarmAnalog[10].FeedPumpTag := 0 ;
   AlarmAnalog[10].TransferPumpEnable := 0 ;
   AlarmAnalog[10].TransferPumpTag := 0 ;
   AlarmAnalog[10].Disable := 0 ;
   AlarmAnalog[10].HIHIEnable := 0 ;
   
   (*AnalogPoint[11]: Filtrate UV AI102
   ============================================================*)
   
   IF Options.No_Device_Connected OR Options.AI101 OR Options.AI101_AI104 THEN
   	AnalogPoint[11].EnableCfg := 0 ;
   	AlarmAnalog[11].EnableCfg := 0 ;
   ELSIF Options.AI102_AI103 OR Options.AI101_AI102_AI103 OR Options.AI101_AI102_AI103_AI104 THEN
   	AnalogPoint[11].EnableCfg := 1 ;
   	AlarmAnalog[11].EnableCfg := 1 ;
   ELSE
   	AnalogPoint[11].EnableCfg := 0 ;
   	AlarmAnalog[11].EnableCfg := 0 ;
   END_IF;
   
   AnalogPoint[11].Address := 11 ;
   AnalogPoint[11].RawMin := 6553 ;
   AnalogPoint[11].RawMax := 32767 ;
   AnalogPoint[11].RealCfg := 1 ;
   AnalogPoint[11].OverrideCfg := 1 ;
   AlarmAnalog[11].FeedPumpEnable := 0 ;
   AlarmAnalog[11].FeedPumpTag := 0 ;
   AlarmAnalog[11].TransferPumpEnable := 0 ;
   AlarmAnalog[11].TransferPumpTag := 0 ;
   AlarmAnalog[11].Disable := 0 ;
   AlarmAnalog[11].HIHIEnable := 0 ;
   
   (*AnalogPoint[12]: Filtrate UV AI103
   ============================================================*)
   
   IF Options.No_Device_Connected OR Options.AI101 OR Options.AI101_AI104 THEN
   	AnalogPoint[12].EnableCfg := 0 ;
   	AlarmAnalog[12].EnableCfg := 0 ;
   ELSIF Options.AI102_AI103 OR Options.AI101_AI102_AI103 OR Options.AI101_AI102_AI103_AI104 THEN
   	AnalogPoint[12].EnableCfg := 1 ;
   	AlarmAnalog[12].EnableCfg := 1 ;
   ELSE
   	AnalogPoint[12].EnableCfg := 0 ;
   	AlarmAnalog[12].EnableCfg := 0 ;
   END_IF;
   
   AnalogPoint[12].Address := 12 ;
   AnalogPoint[12].RawMin := 6553 ;
   AnalogPoint[12].RawMax := 32767 ;
   AnalogPoint[12].RealCfg := 1 ;
   AnalogPoint[12].OverrideCfg := 1 ;
   AlarmAnalog[12].FeedPumpEnable := 0 ;
   AlarmAnalog[12].FeedPumpTag := 0 ;
   AlarmAnalog[12].TransferPumpEnable := 0 ;
   AlarmAnalog[12].TransferPumpTag := 0 ;
   AlarmAnalog[12].Disable := 0 ;
   AlarmAnalog[12].HIHIEnable := 0 ;
   
   (*AnalogPoint[13]: Feed Bag Temperature TI001
   ============================================================*)
   AnalogPoint[13].EnableCfg := 1 ;
   AnalogPoint[13].Address := 13 ;
   AnalogPoint[13].RawMin := 6553 ;
   AnalogPoint[13].RawMax := 32767 ;
   AnalogPoint[13].RealCfg := 1 ;
   AnalogPoint[13].OverrideCfg := 1 ;
   AlarmAnalog[13].FeedPumpEnable := 0 ;
   AlarmAnalog[13].FeedPumpTag := 0 ;
   AlarmAnalog[13].TransferPumpEnable := 0 ;
   AlarmAnalog[13].TransferPumpTag := 0 ;
   AlarmAnalog[13].EnableCfg := 1 ;
   AlarmAnalog[13].Disable := 0 ;
   AlarmAnalog[13].HIHIEnable := 0 ;
   
   (*AnalogPoint[14]: Mixer Speed MIX001
   ============================================================*)
   AnalogPoint[14].EnableCfg := 1 ;
   AnalogPoint[14].Address := 14 ;
   AnalogPoint[14].RawMin := 0 ;
   AnalogPoint[14].RawMax := 16384 ;
   AnalogPoint[14].RealCfg := 1 ;
   AnalogPoint[14].OverrideCfg := 0 ;
   AlarmAnalog[14].FeedPumpEnable := 0 ;
   AlarmAnalog[14].FeedPumpTag := 0 ;
   AlarmAnalog[14].TransferPumpEnable := 0 ;
   AlarmAnalog[14].TransferPumpTag := 0 ;
   AlarmAnalog[14].EnableCfg := 0 ;
   AlarmAnalog[14].Disable := 0 ;
   AlarmAnalog[14].HIHIEnable := 0 ;
   
   (*AnalogPoint[15]: Feed Bag Weight WI001
   ============================================================*)
   AnalogPoint[15].EnableCfg := 1 ;
   AnalogPoint[15].Address := 15 ;
   AnalogPoint[15].RawMin := 0 ;
   AnalogPoint[15].RawMax := 99999 ;
   AnalogPoint[15].RealCfg := 0 ;
   AnalogPoint[15].OverrideCfg := 1 ;
   AnalogPoint[15].ScaledMin := 0 ;
   AnalogPoint[15].ScaledMax := 999.99 ;
   AlarmAnalog[15].FeedPumpEnable := 1 ;
   AlarmAnalog[15].FeedPumpTag := 1 ;
   AlarmAnalog[15].TransferPumpEnable := 0 ;
   AlarmAnalog[15].TransferPumpTag := 0 ;
   AlarmAnalog[15].EnableCfg := 1 ;
   AlarmAnalog[15].Disable := 0 ;
   AlarmAnalog[15].HIHIEnable := 0 ;
   
   (*AnalogPoint[16]: Spare
   ============================================================*)
   AnalogPoint[16].EnableCfg := 0 ;
   AlarmAnalog[16].EnableCfg := 0 ;
   
   (*AnalogPoint[17]: Retentate Flow FI003
   ============================================================*)
   IF Options.FI003 THEN
   	AnalogPoint[17].EnableCfg := 1 ;
   	AlarmAnalog[17].EnableCfg := 1 ;
   ELSE
   	AnalogPoint[17].EnableCfg := 0 ;
   	AlarmAnalog[17].EnableCfg := 0 ;
   END_IF;
   AnalogPoint[17].Address := 17 ;
   AnalogPoint[17].RawMin := 6553 ;
   AnalogPoint[17].RawMax := 32767 ;
   AnalogPoint[17].RealCfg := 1 ;
   AnalogPoint[17].OverrideCfg := 1 ;
   AlarmAnalog[17].FeedPumpEnable := 1 ;
   AlarmAnalog[17].FeedPumpTag := 1 ;
   AlarmAnalog[17].TransferPumpEnable := 1 ;
   AlarmAnalog[17].TransferPumpTag := 2 ;
   AlarmAnalog[17].Disable := 0 ;
   AlarmAnalog[17].HIHIEnable := 0 ;
   
   (*Reset Loop : Set to 0 the AnalogPoint[18 to 39].EnableCfg
   ============================================================*)
   FOR Config.IndexAP := 18 to 39 by 1 do
   	AnalogPoint[Config.IndexAP].EnableCfg := 0 ;
   	AlarmAnalog[Config.IndexAP].EnableCfg := 0 ;
   End_for ;
   
   (*AnalogPoint[40]: Differential Pressure DP
   ============================================================*)
   AnalogPoint[40].EnableCfg := 1 ;
   AnalogPoint[40].Address := 40 ;
   AnalogPoint[40].RawMin := 6553 ;
   AnalogPoint[40].RawMax := 32767 ;
   AnalogPoint[40].RealCfg := 0 ;
   AnalogPoint[40].OverrideCfg := 1 ;
   AlarmAnalog[40].FeedPumpEnable := 1 ;
   AlarmAnalog[40].FeedPumpTag := 1 ;
   AlarmAnalog[40].TransferPumpEnable := 0 ;
   AlarmAnalog[40].TransferPumpTag := 0 ;
   AlarmAnalog[40].EnableCfg := 1 ;
   AlarmAnalog[40].Disable := 0 ;
   AlarmAnalog[40].HIHIEnable := 0 ;
   
   (*AnalogPoint[41]: Trans-Membrane Pressure TMP
   ============================================================*)
   AnalogPoint[41].EnableCfg := 1 ;
   AnalogPoint[41].Address := 41 ;
   AnalogPoint[41].RawMin := 6553 ;
   AnalogPoint[41].RawMax := 32767 ;
   AnalogPoint[41].RealCfg := 0 ;
   AnalogPoint[41].OverrideCfg := 1 ;
   AlarmAnalog[41].FeedPumpEnable := 1 ;
   AlarmAnalog[41].FeedPumpTag := 1 ;
   AlarmAnalog[41].TransferPumpEnable := 0 ;
   AlarmAnalog[41].TransferPumpTag := 0 ;
   AlarmAnalog[41].EnableCfg := 1 ;
   AlarmAnalog[41].Disable := 0 ;
   AlarmAnalog[41].HIHIEnable := 0 ;
   
   (*AnalogPoint[42]: Feed Flow FI001
   ============================================================*)
   AnalogPoint[42].EnableCfg := 1 ;
   AnalogPoint[42].Address := 42 ;
   AnalogPoint[42].RawMin := 6553 ;
   AnalogPoint[42].RawMax := 32767 ;
   AnalogPoint[42].RealCfg := 0 ;
   AnalogPoint[42].OverrideCfg := 1 ;
   AlarmAnalog[42].FeedPumpEnable := 1 ;
   AlarmAnalog[42].FeedPumpTag := 1 ;
   AlarmAnalog[42].TransferPumpEnable := 0 ;
   AlarmAnalog[42].TransferPumpTag := 0 ;
   AlarmAnalog[42].EnableCfg := 1 ;
   AlarmAnalog[42].Disable := 0 ;
   AlarmAnalog[42].HIHIEnable := 0 ;
   
   (*AnalogPoint[43]: Transfer Pump Flow FI401
   ============================================================*)
   AnalogPoint[43].EnableCfg := 1 ;
   AnalogPoint[43].Address := 43 ;
   AnalogPoint[43].RawMin := 6553 ;
   AnalogPoint[43].RawMax := 32767 ;
   AnalogPoint[43].RealCfg := 0 ;
   AnalogPoint[43].OverrideCfg := 1 ;
   AlarmAnalog[43].FeedPumpEnable := 0 ;
   AlarmAnalog[43].FeedPumpTag := 0 ;
   AlarmAnalog[43].TransferPumpEnable := 1 ;
   AlarmAnalog[43].TransferPumpTag := 2 ;
   AlarmAnalog[43].EnableCfg := 1 ;
   AlarmAnalog[43].Disable := 0 ;
   AlarmAnalog[43].HIHIEnable := 0 ;
   
   (*AnalogPoint[44]: Feed Bag Volume LI001
   ============================================================*)
   AnalogPoint[44].EnableCfg := 1 ;
   AnalogPoint[44].Address := 44 ;
   AnalogPoint[44].RawMin := 6553 ;
   AnalogPoint[44].RawMax := 32767 ;
   AnalogPoint[44].RealCfg := 0 ;
   AnalogPoint[44].OverrideCfg := 1 ;
   AlarmAnalog[44].FeedPumpEnable := 1 ;
   AlarmAnalog[44].FeedPumpTag := 1 ;
   AlarmAnalog[44].TransferPumpEnable := 0 ;
   AlarmAnalog[44].TransferPumpTag := 0 ;
   AlarmAnalog[44].EnableCfg := 1 ;
   AlarmAnalog[44].Disable := 0 ;
   AlarmAnalog[44].HIHIEnable := 0 ;
   
   (*AnalogPoint[45]: Normalized Water Permeability NWP
   ============================================================*)
   AnalogPoint[45].EnableCfg := 1 ;
   AnalogPoint[45].Address := 45 ;
   AnalogPoint[45].RawMin := 6553 ;
   AnalogPoint[45].RawMax := 32767 ;
   AnalogPoint[45].RealCfg := 0 ;
   AnalogPoint[45].OverrideCfg := 0 ;
   AlarmAnalog[45].FeedPumpEnable := 0 ;
   AlarmAnalog[45].FeedPumpTag := 0 ;
   AlarmAnalog[45].TransferPumpEnable := 0 ;
   AlarmAnalog[45].TransferPumpTag := 0 ;
   AlarmAnalog[45].EnableCfg := 0 ;
   AlarmAnalog[45].Disable := 0 ;
   AlarmAnalog[45].HIHIEnable := 0 ;
   
   (*AnalogPoint[46]: Membrane Permeability PERM
   ============================================================*)
   AnalogPoint[46].EnableCfg := 1 ;
   AnalogPoint[46].Address := 46 ;
   AnalogPoint[46].RawMin := 6553 ;
   AnalogPoint[46].RawMax := 32767 ;
   AnalogPoint[46].RealCfg := 0 ;
   AnalogPoint[46].OverrideCfg := 0 ;
   AlarmAnalog[46].FeedPumpEnable := 0 ;
   AlarmAnalog[46].FeedPumpTag := 0 ;
   AlarmAnalog[46].TransferPumpEnable := 0 ;
   AlarmAnalog[46].TransferPumpTag := 0 ;
   AlarmAnalog[46].EnableCfg := 0 ;
   AlarmAnalog[46].Disable := 0 ;
   AlarmAnalog[46].HIHIEnable := 0 ;
   
   
   
   (*Reset Loop : Set to 0 the AnalogPoint[45 to 49].EnableCfg
   ============================================================*)
   FOR Config.IndexAP := 47 to 49 by 1 do
   	AnalogPoint[Config.IndexAP].EnableCfg := 0 ;
   	AlarmAnalog[Config.IndexAP].EnableCfg := 0 ;
   End_for ;
END_ROUTINE

ROUTINE Config_ControlLoop   (* structured text *)
   (* =======================================================================
   	Config ControlLoop : Configure ControlLoop Structure
   
   	List of treatments
   		- FIC001 Feed Pump Control Loop
   		- LIC001 Level Control Loop
   		- PCV001 Retentate Control Valve Control Loop
   		- PCV001 Retentate Control Valve Control Loop 5ms
   		- PCV101 Filtrate Control Valve Control Loop
   		- PCV101 Filtrate Control Valve Control Loop 5ms
   		- Reset Loop : Disable unused ControlLoop and Deviation Alarm
   
   -----------------------------------------------------------------------------------------------------------------------------------------------------
   	History
   		2019-AUG-13 - ACTEMIUM - B. Roch - Initial version for Candidate Release 3.00.00.00.a
   		2019-SEP-26 - ACTEMIUM - B. Roch - Initial version for Candidate Release 3.00.00.00.c
   							- add control_loop[3] and control_loop[5] configuration
   =========================================================================*)
   
   (* FIC001 Feed Pump Control Loop
   =========================================================================*)
   (*Index set with ControlLoop number*)
   Config.IndexCL := 1 ;
   (*ControlLoop data structure configuration*)
   ControlLoop[1].LoopCfg := 1 ;
   ControlLoop[1].Auto3 := 0;
   ControlLoop[1].Auto4 := 0;
   ControlLoop[1].RampEnable := 1;
   ControlLoop[1].PIDEnable := 1;
   ControlLoop[1].StepIncrement := 0;
   ControlLoop[1].CycleTime := 0;
   ControlLoop[1].SPAuto3 := 0;
   ControlLoop[1].SPAuto4 := 0;
   ControlLoop[1].RangeMin := 0;
   ControlLoop[1].RangeMax := 100;
   ControlLoop[1].RampTimer.PRE := 3600000;
   ControlLoop[1].PIDTimer.PRE := 250;
   ControlLoop[1].CycleTimer.PRE := 2000;
   ControlLoop[1].DigitalOutput := 0;
   ControlLoop[1].RampCfg := 0;
   ControlLoop[1].Auto1Cfg := 1;
   ControlLoop[1].Auto2Cfg := 1;
   ControlLoop[1].Auto3Cfg := 0;
   ControlLoop[1].Auto4Cfg := 0;
   ControlLoop[1].Auto1PVCfg := 42; //FI001
   ControlLoop[1].Auto2PVCfg := 40; //DP
   ControlLoop[1].Auto3PVCfg := 0;
   ControlLoop[1].Auto4PVCfg := 0;
   ControlLoop[1].Auto1RangeMax := AnalogPoint[42].ScaledMax;
   ControlLoop[1].Auto2RangeMax := AnalogPoint[40].ScaledMax;
   ControlLoop[1].Auto3RangeMax := 0;
   ControlLoop[1].Auto4RangeMax := 0;
   ControlLoop[1].AutoSwitchEnable := 0;
   ControlLoop[1].OutputAddress := 2;
   (*Deviation data structure configuration*)
   AlarmDeviation[1].EnableCfg := 1;
   
   (* LIC001 Level Control Loop
   =========================================================================*)
   (*ControlLoop data structure configuration*)
   ControlLoop[2].LoopCfg := 1 ;
   ControlLoop[2].Auto2 := 0;
   ControlLoop[2].Auto3 := 0;
   ControlLoop[2].Auto4 := 0;
   ControlLoop[2].RampEnable := 1;
   ControlLoop[2].PIDEnable := 1;
   ControlLoop[2].StepIncrement := 0;
   ControlLoop[2].CycleTime := 0;
   ControlLoop[2].SPAuto2 := 0;
   ControlLoop[2].SPAuto3 := 0;
   ControlLoop[2].SPAuto4 := 0;
   ControlLoop[2].RangeMin := 0;
   ControlLoop[2].RangeMax := 100;
   ControlLoop[2].RampTimer.PRE := 3600000;
   ControlLoop[2].PIDTimer.PRE := 250;
   ControlLoop[2].CycleTimer.PRE := 2000;
   ControlLoop[2].DigitalOutput := 0;
   ControlLoop[2].RampCfg := 0;
   ControlLoop[2].Auto1Cfg := 1;
   ControlLoop[2].Auto2Cfg := 0;
   ControlLoop[2].Auto3Cfg := 0;
   ControlLoop[2].Auto4Cfg := 0;
   ControlLoop[2].Auto1PVCfg := 44;
   ControlLoop[2].Auto2PVCfg := 0;
   ControlLoop[2].Auto3PVCfg := 0;
   ControlLoop[2].Auto4PVCfg := 0;
   ControlLoop[2].Auto1RangeMax := AnalogPoint[44].ScaledMax;
   ControlLoop[2].Auto2RangeMax := 0;
   ControlLoop[2].Auto3RangeMax := 0;
   ControlLoop[2].Auto4RangeMax := 0;
   ControlLoop[2].AutoSwitchEnable := 0;
   ControlLoop[2].OutputAddress := 3;
   (*Deviation data structure configuration*)
   AlarmDeviation[2].EnableCfg := 1;
   
   (* PCV001 Retentate Control Valve Control Loop
   =========================================================================*)
   (*ControlLoop data structure configuration*)
   ControlLoop[3].LoopCfg := 1 ;
   ControlLoop[3].Auto3 := 0;
   ControlLoop[3].Auto4 := 0;
   ControlLoop[3].PIDEnable := 1;
   ControlLoop[3].StepIncrement := 0;
   ControlLoop[3].CycleTime := 0;
   ControlLoop[3].SPAuto3 := 0;
   ControlLoop[3].SPAuto4 := 0;
   ControlLoop[3].RangeMin := 0;
   ControlLoop[3].RangeMax := 100;
   ControlLoop[3].RampTimer.PRE := 3600000;
   ControlLoop[3].PIDTimer.PRE := 250;
   ControlLoop[3].CycleTimer.PRE := 2000;
   ControlLoop[3].On := 0;
   ControlLoop[3].DigitalOutput := 0;
   ControlLoop[3].RampCfg := 0;
   ControlLoop[3].Auto1Cfg := 1;
   ControlLoop[3].Auto2Cfg := 1;
   ControlLoop[3].Auto3Cfg := 0;
   ControlLoop[3].Auto4Cfg := 0;
   ControlLoop[3].Auto1PVCfg := 6; //PI002
   ControlLoop[3].Auto2PVCfg := 41; //TMP
   ControlLoop[3].Auto3PVCfg := 0;
   ControlLoop[3].Auto4PVCfg := 0;
   ControlLoop[3].Auto1RangeMax := AnalogPoint[6].ScaledMax;
   ControlLoop[3].Auto2RangeMax := AnalogPoint[41].ScaledMax;
   ControlLoop[3].Auto3RangeMax := 0;
   ControlLoop[3].Auto4RangeMax := 0;
   ControlLoop[3].AutoSwitchEnable := 0;
   ControlLoop[3].OutputAddress := 0;
   (*Deviation data structure configuration*)
   AlarmDeviation[3].EnableCfg := 1;
   (*PCV Control : 0-100 %Clo*)
   PCV001_Control.FullOpenSP := 0 ;
   PCV001_Control.FullCloseSP := 100 ;
   PCV001_Control.FullOpenResetTimer.PRE := 1000 ;
   PCV001_Control.FullCloseResetTimer.PRE := 1000 ;
   
   (* PCV001 Retentate Control Valve Control Loop 5ms
   =========================================================================*)
   (*ControlLoop data structure configuration*)
   ControlLoop[4].LoopCfg := 0 ;
   ControlLoop[4].Manual := 0;
   ControlLoop[4].Auto1 := 0;
   ControlLoop[4].Auto2 := 0;
   ControlLoop[4].Auto3 := 0;
   ControlLoop[4].Auto4 := 0;
   ControlLoop[4].PIDEnable := 1;
   ControlLoop[4].RampEnable := 0;
   ControlLoop[4].StepIncrement := 0;
   ControlLoop[4].CycleTime := 0;
   ControlLoop[4].SPAuto1 := 0;
   ControlLoop[4].SPAuto2 := 0;
   ControlLoop[4].SPAuto3 := 0;
   ControlLoop[4].SPAuto4 := 0;
   ControlLoop[4].RangeMin := 0;
   ControlLoop[4].RangeMax := 100;
   ControlLoop[4].RampTimer.PRE := 3600000;
   ControlLoop[4].PIDTimer.PRE := 250;
   ControlLoop[4].CycleTimer.PRE := 2000;
   ControlLoop[4].On := 0;
   ControlLoop[4].DigitalOutput := 0;
   ControlLoop[4].RampCfg := 0;
   ControlLoop[4].Auto1Cfg := 0;
   ControlLoop[4].Auto2Cfg := 0;
   ControlLoop[4].Auto3Cfg := 0;
   ControlLoop[4].Auto4Cfg := 0;
   ControlLoop[4].Auto1PVCfg := 0;
   ControlLoop[4].Auto2PVCfg := 0;
   ControlLoop[4].Auto3PVCfg := 0;
   ControlLoop[4].Auto4PVCfg := 0;
   ControlLoop[4].Auto1RangeMax := 0;
   ControlLoop[4].Auto2RangeMax := 0;
   ControlLoop[4].Auto3RangeMax := 0;
   ControlLoop[4].Auto4RangeMax := 0;
   ControlLoop[4].AutoSwitchEnable := 0;
   ControlLoop[4].OutputAddress := 0;
   ControlLoop[4].PID.KP := 0.2;
   ControlLoop[4].PID.KD := 0.01;
   ControlLoop[4].PID.DB := 0.3;
   ControlLoop[4].PID.UPD := 0.005;
   ControlLoop[4].PID.MAXS := 100;
   ControlLoop[4].PID.MAXO := 100;
   ControlLoop[4].PID.MAXI := 100;
   ControlLoop[4].PID.MAXCV := 100;
   ControlLoop[4].PID.MAXTIE := 4095;
   
   (* PCV101 Filtrate Control Valve Control Loop
   =========================================================================*)
   
   (*If no filtrate measurement disable the flow control mode*)
   IF Options.No_Filtrate_Measurement THEN
   	ControlLoop[5].Auto1 := 0;
   	ControlLoop[5].Auto1Cfg := 0;
   ELSE
   	ControlLoop[5].Auto1Cfg := 1;
   END_IF;
   
   (*ControlLoop data structure configuration*)
   ControlLoop[5].LoopCfg := 1 ;
   ControlLoop[5].Auto3 := 0;
   ControlLoop[5].Auto4 := 0;
   ControlLoop[5].PIDEnable := 1;
   ControlLoop[5].StepIncrement := 0;
   ControlLoop[5].CycleTime := 0;
   ControlLoop[5].SPAuto3 := 0;
   ControlLoop[5].SPAuto4 := 0;
   ControlLoop[5].RangeMin := 0;
   ControlLoop[5].RangeMax := 100;
   ControlLoop[5].RampTimer.PRE := 3600000;
   ControlLoop[5].PIDTimer.PRE := 250;
   ControlLoop[5].CycleTimer.PRE := 2000;
   ControlLoop[5].On := 0;
   ControlLoop[5].DigitalOutput := 0;
   ControlLoop[5].RampCfg := 0;
   ControlLoop[5].Auto2Cfg := 1;
   ControlLoop[5].Auto3Cfg := 0;
   ControlLoop[5].Auto4Cfg := 0;
   ControlLoop[5].Auto1PVCfg := 2; // FI101
   ControlLoop[5].Auto2PVCfg := 41; // TMP
   ControlLoop[5].Auto3PVCfg := 0;
   ControlLoop[5].Auto4PVCfg := 0;
   ControlLoop[5].Auto1RangeMax := AnalogPoint[2].ScaledMax;
   ControlLoop[5].Auto2RangeMax := AnalogPoint[41].ScaledMax;
   ControlLoop[5].Auto3RangeMax := 0;
   ControlLoop[5].Auto4RangeMax := 0;
   ControlLoop[5].AutoSwitchEnable := 0;
   ControlLoop[5].OutputAddress := 1;
   (*Deviation data structure configuration*)
   AlarmDeviation[5].EnableCfg := 1;
   (*PCV Control : 0-100 %opn*)
   PCV101_Control.FullOpenSP := 100 ;
   PCV101_Control.FullCloseSP := 0 ;
   PCV101_Control.FullOpenResetTimer.PRE := 1000 ;
   PCV101_Control.FullCloseResetTimer.PRE := 1000 ;
   
   
   (* PCV101 Filtrate Control Valve Control Loop
   =========================================================================*)
   
   (*ControlLoop data structure configuration*)
   ControlLoop[6].LoopCfg := 0 ;
   ControlLoop[6].Manual := 0;
   ControlLoop[6].Auto1 := 0;
   ControlLoop[6].Auto2 := 0;
   ControlLoop[6].Auto3 := 0;
   ControlLoop[6].Auto4 := 0;
   ControlLoop[6].PIDEnable := 1;
   ControlLoop[6].RampEnable := 0;
   ControlLoop[6].StepIncrement := 0;
   ControlLoop[6].CycleTime := 0;
   ControlLoop[6].SPAuto1 := 0;
   ControlLoop[6].SPAuto2 := 0;
   ControlLoop[6].SPAuto3 := 0;
   ControlLoop[6].SPAuto4 := 0;
   ControlLoop[6].RangeMin := 0;
   ControlLoop[6].RangeMax := 100;
   ControlLoop[6].RampTimer.PRE := 3600000;
   ControlLoop[6].PIDTimer.PRE := 250;
   ControlLoop[6].CycleTimer.PRE := 2000;
   ControlLoop[6].On := 0;
   ControlLoop[6].DigitalOutput := 0;
   ControlLoop[6].RampCfg := 0;
   ControlLoop[6].Auto1Cfg := 0;
   ControlLoop[6].Auto2Cfg := 0;
   ControlLoop[6].Auto3Cfg := 0;
   ControlLoop[6].Auto4Cfg := 0;
   ControlLoop[6].Auto1PVCfg := 0;
   ControlLoop[6].Auto2PVCfg := 0;
   ControlLoop[6].Auto3PVCfg := 0;
   ControlLoop[6].Auto4PVCfg := 0;
   ControlLoop[6].Auto1RangeMax := 0;
   ControlLoop[6].Auto2RangeMax := 0;
   ControlLoop[6].Auto3RangeMax := 0;
   ControlLoop[6].Auto4RangeMax := 0;
   ControlLoop[6].AutoSwitchEnable := 0;
   ControlLoop[6].OutputAddress := 1;
   ControlLoop[6].PID.KP := 0.3;
   ControlLoop[6].PID.KD := 0.01;
   ControlLoop[6].PID.DB := 0.3;
   ControlLoop[6].PID.UPD := 0.005;
   ControlLoop[6].PID.MAXS := 100;
   ControlLoop[6].PID.MAXO := 100;
   ControlLoop[6].PID.MAXI := 100;
   ControlLoop[6].PID.MAXCV := 100;
   ControlLoop[6].PID.MAXTIE := 4095;
   
   (*Reset Loop : Disable unused ControlLoop and Deviation Alarm
   ============================================================*)
   ControlLoop[0].LoopCfg := 0 ;
   AlarmDeviation[0].EnableCfg := 0;
   AlarmDeviation[0].Override := 1;
   AlarmDeviation[0].Disable := 1;
   ControlLoop[4].LoopCfg := 0 ;
   AlarmDeviation[4].EnableCfg := 0;
   AlarmDeviation[4].Override := 1;
   AlarmDeviation[4].Disable := 1;
   ControlLoop[6].LoopCfg := 0 ;
   AlarmDeviation[6].EnableCfg := 0;
   AlarmDeviation[6].Override := 1;
   AlarmDeviation[6].Disable := 1;
   
   FOR Config.IndexCL := 7 to 19 do
   	ControlLoop[Config.IndexCL].LoopCfg := 0 ;
   	AlarmDeviation[Config.IndexCL].EnableCfg := 0;
   	AlarmDeviation[Config.IndexCL].Override := 1;
   	AlarmDeviation[Config.IndexCL].Disable := 1;
   End_for ;
END_ROUTINE

ROUTINE Config_DigitalPoint_Real   (* structured text *)
// Apply the default configuration
   (* ==========================================================
   	Config DigitalPoint Real : Configure DigitalPoint Structure (for real input)
   
   	List of treatments
   		- DigitalPoint[0] : Valves Air Defect PSL602
   		- DigitalPoint[1] : Door Closed XS001
   		- DigitalPoint[2] : Door to Frame Locking Closed XS006
   		- DigitalPoint[3] : Emergency Stop ES001
   		- DigitalPoint[4] : Feed Pump High Pressure PSH001
   		- DigitalPoint[5] : Transfer Pump High Pressure PSH401
   		- DigitalPoint[6] : Clamshell Locking 1 Closed XS002
   		- DigitalPoint[7] : Clamshell Locking 2 Closed XS003
   		- DigitalPoint[8] : Feed Pump Defect SIC001DF
   		- DigitalPoint[9] : Transfer Pump Defect SIC002DF
   		- DigitalPoint[10]: Manifold Valves Air Defect PSL603
   		- DigitalPoint[11]: Pump P001 Type XS011
   		- DigitalPoint[12]: Pump P002 Type XS012
   		- DigitalPoint[13]: C8000 Defect XC102_3DF
   		- DigitalPoint[14]: Mixer Defect SIC003DF
   		- DigitalPoint[15]: Tank Skid Remote / Standalone SRL001
   		- Reset Loop : Set to 0 the DigitalPoint[16 to 49].EnableCfg
   
   -----------------------------------------------------------------------------------------------------------------------------------------------------
   	History
   		2019-AUG-13 - ACTEMIUM - B. Roch - Initial version for Candidate Release 3.00.00.00.a
   		2020-SEP-21 - Merck - Q. Spindler - Modifications for Candidate Release 3.00.00.01.a
   							- Reset XS011 and XS012 currentvalue if the MoldType is not 123
   ============================================================*)
   
   (*DigitalPoint[0] : Valves Air Defect PSL602
   ============================================================*)
   DigitalPoint[0].EnableCfg := 1 ;
   DigitalPoint[0].ActiveStateCFg := 1 ;
   DigitalPoint[0].RealInputCfg := 1 ;
   DigitalPoint[0].InputAddressCfg := 0 ;
   DigitalPoint[0].AlarmCfg := 1 ;
   DigitalPoint[0].AlarmStateCfg := 0 ;
   DigitalPoint[0].OverrideCfg := 1 ;
   DigitalPoint[0].PriorityCfg := 1 ;
   DigitalPoint[0].Cond1Cfg := 0 ;
   DigitalPoint[0].Cond2Cfg := 0 ;
   DigitalPoint[0].FlashingInputCfg := 0 ;
   
   (*DigitalPoint[1] : Door Closed XS001
   ============================================================*)
   DigitalPoint[1].EnableCfg := 1 ;
   DigitalPoint[1].ActiveStateCFg := 1 ;
   DigitalPoint[1].RealInputCfg := 1 ;
   DigitalPoint[1].InputAddressCfg := 1 ;
   DigitalPoint[1].AlarmCfg := 1 ;
   DigitalPoint[1].AlarmStateCfg := 0 ;
   DigitalPoint[1].OverrideCfg := 1 ;
   DigitalPoint[1].PriorityCfg := 0 ;
   DigitalPoint[1].Priority := 1 ;
   DigitalPoint[1].Cond1Cfg := 0 ;
   DigitalPoint[1].Cond2Cfg := 0 ;
   DigitalPoint[1].FlashingInputCfg := 0 ;
   
   (*DigitalPoint[2] : Door to Frame Locking Closed XS006
   ============================================================*)
   DigitalPoint[2].EnableCfg := 1 ;
   DigitalPoint[2].ActiveStateCFg := 1 ;
   DigitalPoint[2].RealInputCfg := 1 ;
   DigitalPoint[2].InputAddressCfg := 2 ;
   DigitalPoint[2].AlarmCfg := 0 ;
   DigitalPoint[2].AlarmStateCfg := 0 ;
   DigitalPoint[2].OverrideCfg := 0 ;
   DigitalPoint[2].PriorityCfg := 0 ;
   DigitalPoint[2].Cond1Cfg := 0 ;
   DigitalPoint[2].Cond2Cfg := 0 ;
   DigitalPoint[2].FlashingInputCfg := 0 ;
   
   (*DigitalPoint[3] : Emergency Stop ES001
   ============================================================*)
   DigitalPoint[3].EnableCfg := 1 ;
   DigitalPoint[3].ActiveStateCFg := 1 ;
   DigitalPoint[3].RealInputCfg := 1 ;
   DigitalPoint[3].InputAddressCfg := 3 ;
   DigitalPoint[3].AlarmCfg := 1 ;
   DigitalPoint[3].AlarmStateCfg := 0 ;
   DigitalPoint[3].OverrideCfg := 0 ;
   DigitalPoint[3].Priority := 1 ;
   DigitalPoint[3].PriorityCfg := 0 ;
   DigitalPoint[3].Cond1Cfg := 0 ;
   DigitalPoint[3].Cond2Cfg := 0 ;
   DigitalPoint[3].FlashingInputCfg := 0 ;
   
   (*DigitalPoint[4] : Feed Pump High Pressure PSH001
   ============================================================*)
   DigitalPoint[4].EnableCfg := 1 ;
   DigitalPoint[4].ActiveStateCFg := 1 ;
   DigitalPoint[4].RealInputCfg := 1 ;
   DigitalPoint[4].InputAddressCfg := 4 ;
   DigitalPoint[4].AlarmCfg := 1 ;
   DigitalPoint[4].AlarmStateCfg := 0 ;
   DigitalPoint[4].OverrideCfg := 1 ;
   DigitalPoint[4].PriorityCfg := 0 ;
   DigitalPoint[4].Priority := 1 ;
   DigitalPoint[4].Cond1Cfg := 0 ;
   DigitalPoint[4].Cond2Cfg := 0 ;
   DigitalPoint[4].FlashingInputCfg := 0 ;
   
   (*DigitalPoint[5] : Transfer Pump High Pressure PSH401
   ============================================================*)
   DigitalPoint[5].EnableCfg := 1 ;
   DigitalPoint[5].ActiveStateCFg := 1 ;
   DigitalPoint[5].RealInputCfg := 1 ;
   DigitalPoint[5].InputAddressCfg := 5 ;
   DigitalPoint[5].AlarmCfg := 1 ;
   DigitalPoint[5].AlarmStateCfg := 0 ;
   DigitalPoint[5].OverrideCfg := 1 ;
   DigitalPoint[5].PriorityCfg := 0 ;
   DigitalPoint[5].Priority := 1 ;
   DigitalPoint[5].Cond1Cfg := 0 ;
   DigitalPoint[5].Cond2Cfg := 0 ;
   DigitalPoint[5].FlashingInputCfg := 0 ;
   
   (*DigitalPoint[6] : Clamshell Locking 1 Closed XS002
   ============================================================*)
   DigitalPoint[6].EnableCfg := 1 ;
   DigitalPoint[6].ActiveStateCFg := 1 ;
   DigitalPoint[6].RealInputCfg := 1 ;
   DigitalPoint[6].InputAddressCfg := 6 ;
   DigitalPoint[6].AlarmCfg := 0 ;
   DigitalPoint[6].AlarmStateCfg := 0 ;
   DigitalPoint[6].OverrideCfg := 0 ;
   DigitalPoint[6].PriorityCfg := 0 ;
   DigitalPoint[6].Cond1Cfg := 0 ;
   DigitalPoint[6].Cond2Cfg := 0 ;
   DigitalPoint[6].FlashingInputCfg := 0 ;
   
   (*DigitalPoint[7] : Clamshell Locking 2 Closed XS003
   ============================================================*)
   DigitalPoint[7].EnableCfg := 1 ;
   DigitalPoint[7].ActiveStateCFg := 1 ;
   DigitalPoint[7].RealInputCfg := 1 ;
   DigitalPoint[7].InputAddressCfg := 7 ;
   DigitalPoint[7].AlarmCfg := 0 ;
   DigitalPoint[7].AlarmStateCfg := 0 ;
   DigitalPoint[7].OverrideCfg := 0 ;
   DigitalPoint[7].PriorityCfg := 0 ;
   DigitalPoint[7].Cond1Cfg := 0 ;
   DigitalPoint[7].Cond2Cfg := 0 ;
   DigitalPoint[7].FlashingInputCfg := 0 ;
   
   (*DigitalPoint[8] : Feed Pump Defect SIC001DF
   ============================================================*)
   DigitalPoint[8].EnableCfg := 1 ;
   DigitalPoint[8].ActiveStateCFg := 1 ;
   DigitalPoint[8].RealInputCfg := 1 ;
   DigitalPoint[8].InputAddressCfg := 8 ;
   DigitalPoint[8].AlarmCfg := 1 ;
   DigitalPoint[8].AlarmStateCfg := 0 ;
   DigitalPoint[8].OverrideCfg := 1 ;
   DigitalPoint[8].PriorityCfg := 1 ;
   DigitalPoint[8].Cond1Cfg := 0 ;
   DigitalPoint[8].Cond2Cfg := 0 ;
   DigitalPoint[8].FlashingInputCfg := 0 ;
   
   (*DigitalPoint[9] : Transfer Pump Defect SIC002DF
   ============================================================*)
   DigitalPoint[9].EnableCfg := 1 ;
   DigitalPoint[9].ActiveStateCFg := 1 ;
   DigitalPoint[9].RealInputCfg := 1 ;
   DigitalPoint[9].InputAddressCfg := 9 ;
   DigitalPoint[9].AlarmCfg := 1 ;
   DigitalPoint[9].AlarmStateCfg := 0 ;
   DigitalPoint[9].OverrideCfg := 1 ;
   DigitalPoint[9].PriorityCfg := 1 ;
   DigitalPoint[9].Cond1Cfg := 0 ;
   DigitalPoint[9].Cond2Cfg := 0 ;
   DigitalPoint[9].FlashingInputCfg := 0 ;
   
   (*DigitalPoint[10]: Manifold Valves Air Defect PSL603
   ============================================================*)
   DigitalPoint[10].EnableCfg := 1 ;
   DigitalPoint[10].ActiveStateCFg := 1 ;
   DigitalPoint[10].RealInputCfg := 1 ;
   DigitalPoint[10].InputAddressCfg := 10 ;
   DigitalPoint[10].AlarmCfg := 1 ;
   DigitalPoint[10].AlarmStateCfg := 0 ;
   DigitalPoint[10].OverrideCfg := 1 ;
   DigitalPoint[10].PriorityCfg := 1 ;
   DigitalPoint[10].Cond1Cfg := 0 ;
   DigitalPoint[10].Cond2Cfg := 0 ;
   DigitalPoint[10].FlashingInputCfg := 0 ;
   
   (*DigitalPoint[11]: Pump P001 Type XS011
   ============================================================*)
   
   IF ThisSystem.MoldType = 123 THEN
   	DigitalPoint[11].EnableCfg := 1 ;
   ELSIF ThisSystem.MoldType = 124 THEN
   	DigitalPoint[11].EnableCfg := 0 ;
   	DigitalPoint[11].CurrentValue := 0 ;
   ELSE
   	DigitalPoint[11].EnableCfg := 0 ;
   	DigitalPoint[11].CurrentValue := 0 ;
   END_IF;
   
   DigitalPoint[11].ActiveStateCFg := 1 ;
   DigitalPoint[11].RealInputCfg := 1 ;
   DigitalPoint[11].InputAddressCfg := 11 ;
   DigitalPoint[11].AlarmCfg := 0 ;
   DigitalPoint[11].AlarmStateCfg := 0 ;
   DigitalPoint[11].OverrideCfg := 0 ;
   DigitalPoint[11].PriorityCfg := 0 ;
   DigitalPoint[11].Cond1Cfg := 0 ;
   DigitalPoint[11].Cond2Cfg := 0 ;
   DigitalPoint[11].FlashingInputCfg := 0 ;
   
   (*DigitalPoint[12]: Pump P002 Type XS012
   ============================================================*)
   
   IF ThisSystem.MoldType = 123 THEN
   	DigitalPoint[12].EnableCfg := 1 ;
   ELSIF ThisSystem.MoldType = 124 THEN
   	DigitalPoint[12].EnableCfg := 0 ;
   	DigitalPoint[12].CurrentValue := 0 ;
   ELSE
   	DigitalPoint[12].EnableCfg := 0 ;
   	DigitalPoint[12].CurrentValue := 0 ;
   END_IF;
   
   DigitalPoint[12].EnableCfg := 1 ;
   DigitalPoint[12].ActiveStateCFg := 1 ;
   DigitalPoint[12].RealInputCfg := 1 ;
   DigitalPoint[12].InputAddressCfg := 12 ;
   DigitalPoint[12].AlarmCfg := 0 ;
   DigitalPoint[12].AlarmStateCfg := 0 ;
   DigitalPoint[12].OverrideCfg := 0 ;
   DigitalPoint[12].PriorityCfg := 0 ;
   DigitalPoint[12].Cond1Cfg := 0 ;
   DigitalPoint[12].Cond2Cfg := 0 ;
   DigitalPoint[12].FlashingInputCfg := 0 ;
   
   (*DigitalPoint[13]: C8000 Defect XC102_3DF
   ============================================================*)
   
   IF Options.No_Device_Connected OR Options.AI101 OR Options.AI101_AI104 THEN
   	DigitalPoint[13].EnableCfg := 0 ;
   	DigitalPoint[13].AlarmCfg := 0 ;
   	DigitalPoint[13].Alarm := 0 ;
   ELSIF Options.AI102_AI103 OR Options.AI101_AI102_AI103 OR Options.AI101_AI102_AI103_AI104 THEN
   	DigitalPoint[13].EnableCfg := 1 ;
   	DigitalPoint[13].AlarmCfg := 1 ;
   ELSE
   	DigitalPoint[13].EnableCfg := 0 ;
   	DigitalPoint[13].AlarmCfg := 0 ;
   	DigitalPoint[13].Alarm := 0 ;
   END_IF;
   
   DigitalPoint[13].ActiveStateCFg := 1 ;
   DigitalPoint[13].RealInputCfg := 1 ;
   DigitalPoint[13].InputAddressCfg := 13 ;
   DigitalPoint[13].AlarmStateCfg := 0 ;
   DigitalPoint[13].OverrideCfg := 1 ;
   DigitalPoint[13].PriorityCfg := 1 ;
   DigitalPoint[13].Cond1Cfg := 0 ;
   DigitalPoint[13].Cond2Cfg := 0 ;
   DigitalPoint[13].FlashingInputCfg := 0 ;
   
   (*DigitalPoint[14]: Mixer Defect SIC003DF
   ============================================================*)
   DigitalPoint[14].EnableCfg := 1 ;
   DigitalPoint[14].ActiveStateCFg := 1 ;
   DigitalPoint[14].RealInputCfg := 1 ;
   DigitalPoint[14].InputAddressCfg := 14 ;
   DigitalPoint[14].AlarmCfg := 1 ;
   DigitalPoint[14].AlarmStateCfg := 0 ;
   DigitalPoint[14].OverrideCfg := 1 ;
   DigitalPoint[14].PriorityCfg := 1 ;
   DigitalPoint[14].Cond1Cfg := 0 ;
   DigitalPoint[14].Cond2Cfg := 0 ;
   DigitalPoint[14].FlashingInputCfg := 0 ;
   
   (*DigitalPoint[15]: Tank Skid Remote / Standalone SRL001
   ============================================================*)
   DigitalPoint[15].EnableCfg := 1 ;
   DigitalPoint[15].ActiveStateCFg := 1 ;
   DigitalPoint[15].RealInputCfg := 1 ;
   DigitalPoint[15].InputAddressCfg := 15 ;
   DigitalPoint[15].AlarmCfg := 0 ;
   DigitalPoint[15].AlarmStateCfg := 0 ;
   DigitalPoint[15].OverrideCfg := 0 ;
   DigitalPoint[15].PriorityCfg := 0 ;
   DigitalPoint[15].Cond1Cfg := 0 ;
   DigitalPoint[15].Cond2Cfg := 0 ;
   DigitalPoint[15].FlashingInputCfg := 0 ;
   
   
   
   (*Reset Loop : Set to 0 the DigitalPoint[16 to 49].EnableCfg
   ============================================================*)
   FOR Config.IndexDP := 16 to 49 do
   	DigitalPoint[Config.IndexDP].EnableCfg := 0 ;
   	DigitalPoint[Config.IndexDP].AlarmCfg := 0 ;
   End_for ;
END_ROUTINE

ROUTINE Config_DigitalPoint_Soft   (* structured text *)
   (* ==========================================================
   	Config DigitalPoint Soft : Configure DigitalPoint Structure (for soft input)
   
   	List of treatments
   		- DigitalPoint[50]: YA01 PC to PLC Com. Failure
   		- DigitalPoint[51]: YA02 CCP Runtime Com. Failure
   		- DigitalPoint[52]: YA03 Historical Data Collection Failure
   		- DigitalPoint[53]: YA04 Hard drive Overload
   		- DigitalPoint[54]: YA05 Database Overload
   		- DigitalPoint[55]: YA06 Node 0 Communication Failure - Smart
   		- DigitalPoint[56]: YA07 Node 0 Internal Defect - Smart
   		- DigitalPoint[57]: YA08 Node 1 Communication Failure - Clamshell
   		- DigitalPoint[58]: YA09 Node 1 Internal Defect - Clamshell
   		- DigitalPoint[59]: YA10 PLC Program Major Fault
   		- DigitalPoint[60]: YA11 Database Corrupted
   		- DigitalPoint[61]: YA12 Unauthorized accesses
   		- DigitalPoint[62]: YA13 Tank Size Mismatch
   		- DigitalPoint[63]: YA14 SQL Server Write Failure
   		- DigitalPoint[64]: UserNCr1 User Non Critical Alarm 1
   		- DigitalPoint[65]: UserCr1 User Critical Alarm 1
   		- DigitalPoint[66]: UserNCr2 User Non Critical Alarm 2
   		- DigitalPoint[67]: UserCr2 User Critical Alarm 2
   		- DigitalPoint[68]: ZSDF Clamshell Locking Defect
   		- DigitalPoint[69]: YA15 Node 3 Communication Failure - Pump
   		- DigitalPoint[70]: YA16 Node 3 Internal Defect - Pump
   		- DigitalPoint[71]: YA17 Node 4 Communication Failure - Instrum
   		- DigitalPoint[72]: YA18 Node 4 Internal Defect - Instrum
   		- DigitalPoint[73]: YA19 Node 5 Communication Failure - Tank
   		- DigitalPoint[74]: YA20 Node 5 Internal Defect - Tank
   		- DigitalPoint[75]: YA21 IND331 Communication Failure
   		- DigitalPoint[76]: YA22 IND131 Communication Failure
   		- DigitalPoint[77]: YA41 Operating Time Exceeded
   		- Reset Loop : Set to 0 the DigitalPoint[77 to 89].EnableCfg
   		- DigitalPoint[90]: AI101_SIG Filtrate Conductivity Signal default
   		- DigitalPoint[91]: AI102_SIG Filtrate UV Signal default
   		- DigitalPoint[92]: AI103_SIG Filtrate UV Signal default
   		- DigitalPoint[93]: FI101_SIG Filtrate Flow flow Signal default
   		- DigitalPoint[94]: WI001_SIG Feed Bag Weight Signal default
   		- DigitalPoint[95]: WI101_SIG Filtrate Weight Signal default
   		- DigitalPoint[96]: WI102_SIG Customer Filtrate Weight Signal default
   		- DigitalPoint[97]: PI001_SIG Feed Pressure Signal default
   		- DigitalPoint[98]: PI002_SIG Retentate Pressure Signal default
   		- DigitalPoint[99]: PI101_SIG Filtrate Pressure Signal default
   		- DigitalPoint[100]: PI401_SIG Transfer Pump Pressure Signal default
   		- DigitalPoint[101]: TI001_SIG Feed Bag Temperature Signal default
   		- DigitalPoint[102]: PCV001_SIG PCV001 Position Signal default
   		- DigitalPoint[103]: PCV101_SIG PCV101 Position Signal default
   		- DigitalPoint[104]: MIX001_SIG Mixer Speed Signal default
   		- DigitalPoint[105]: AI104_SIG Filtrate pH Signal default
   		- DigitalPoint[106]: FI003_SIG Retentate Flow Signal default
   		- Reset Loop : Set to 0 the DigitalPoint[107 to 149].EnableCfg
   
   -----------------------------------------------------------------------------------------------------------------------------------------------------
   	History
   		2019-AUG-13 - ACTEMIUM - B. Roch - Initial version for Candidate Release 3.00.00.00.a
   		2020-SEP-29 - Merck - Q. Spindler - Modifications for Candidate Release 3.00.00.01.a
   					- Add FI003_SIG
   		2020-NOV-23 - Merck - Q. Spindler - Modifications for Candidate Release 3.00.00.01.b
   					- Remove force of ZSDF priority
   					- Change FI003_SIG option
   		2021-APR-27 - DAVIDSON- Ch. ARBOGAST - Modifications for Candidate Release 3.01.00.00.a
   					- add DigitalPoint[77]: YA41 Operating Time Exceeded
   ============================================================*)
   
   (*DigitalPoint[50]: YA01 PC to PLC Com. Failure
   ============================================================*)
   DigitalPoint[50].EnableCfg := 1 ;
   DigitalPoint[50].ActiveStateCFg := 0 ;
   DigitalPoint[50].RealInputCfg := 0 ;
   DigitalPoint[50].InputAddressCfg := 50 ;
   DigitalPoint[50].AlarmCfg := 1 ;
   DigitalPoint[50].AlarmStateCfg := 1 ;
   DigitalPoint[50].OverrideCfg := 1 ;
   DigitalPoint[50].PriorityCfg := 1 ;
   DigitalPoint[50].Cond1Cfg := 1 ;
   DigitalPoint[50].Cond2Cfg := 0 ;
   DigitalPoint[50].FlashingInputCfg := 0 ;
   
   (*DigitalPoint[51]: YA02 CCP Runtime Com. Failure
   ============================================================*)
   DigitalPoint[51].EnableCfg := 1 ;
   DigitalPoint[51].ActiveStateCFg := 0 ;
   DigitalPoint[51].RealInputCfg := 0 ;
   DigitalPoint[51].InputAddressCfg := 51 ;
   DigitalPoint[51].AlarmCfg := 1 ;
   DigitalPoint[51].AlarmStateCfg := 1 ;
   DigitalPoint[51].OverrideCfg := 1 ;
   DigitalPoint[51].PriorityCfg := 1 ;
   DigitalPoint[51].Cond1Cfg := 1 ;
   DigitalPoint[51].Cond2Cfg := 0 ;
   DigitalPoint[51].FlashingInputCfg := 0 ;
   
   (*DigitalPoint[52]: YA03 Historical Data Collection Failure
   ============================================================*)
   DigitalPoint[52].EnableCfg := 1 ;
   DigitalPoint[52].ActiveStateCFg := 0 ;
   DigitalPoint[52].RealInputCfg := 0 ;
   DigitalPoint[52].InputAddressCfg := 52 ;
   DigitalPoint[52].AlarmCfg := 1 ;
   DigitalPoint[52].AlarmStateCfg := 1 ;
   DigitalPoint[52].OverrideCfg := 1 ;
   DigitalPoint[52].PriorityCfg := 1 ;
   DigitalPoint[52].Cond1Cfg := 1 ;
   DigitalPoint[52].Cond2Cfg := 0 ;
   DigitalPoint[52].FlashingInputCfg := 0 ;
   
   (*DigitalPoint[53]: YA04 Hard drive Overload
   ============================================================*)
   DigitalPoint[53].EnableCfg := 1 ;
   DigitalPoint[53].ActiveStateCFg := 1 ;
   DigitalPoint[53].RealInputCfg := 0 ;
   DigitalPoint[53].InputAddressCfg := 53 ;
   DigitalPoint[53].AlarmCfg := 1 ;
   DigitalPoint[53].AlarmStateCfg := 1 ;
   DigitalPoint[53].OverrideCfg := 1 ;
   DigitalPoint[53].PriorityCfg := 1 ;
   DigitalPoint[53].Cond1Cfg := 0 ;
   DigitalPoint[53].Cond2Cfg := 0 ;
   DigitalPoint[53].FlashingInputCfg := 0 ;
   
   (*DigitalPoint[54]: YA05 Database Overload
   ============================================================*)
   DigitalPoint[54].EnableCfg := 1 ;
   DigitalPoint[54].ActiveStateCFg := 1 ;
   DigitalPoint[54].RealInputCfg := 0 ;
   DigitalPoint[54].InputAddressCfg := 54 ;
   DigitalPoint[54].AlarmCfg := 1 ;
   DigitalPoint[54].AlarmStateCfg := 1 ;
   DigitalPoint[54].OverrideCfg := 1 ;
   DigitalPoint[54].PriorityCfg := 1 ;
   DigitalPoint[54].Cond1Cfg := 0 ;
   DigitalPoint[54].Cond2Cfg := 0 ;
   DigitalPoint[54].FlashingInputCfg := 0 ;
   
   (*DigitalPoint[55]: YA06 Node 0 Communication Failure - Smart
   ============================================================*)
   DigitalPoint[55].EnableCfg := 1 ;
   DigitalPoint[55].ActiveStateCFg := 1 ;
   DigitalPoint[55].RealInputCfg := 0;
   DigitalPoint[55].InputAddressCfg := 55 ;
   DigitalPoint[55].AlarmCfg := 1 ;
   DigitalPoint[55].AlarmStateCfg := 1 ;
   DigitalPoint[55].OverrideCfg := 1 ;
   DigitalPoint[55].PriorityCfg := 1 ;
   DigitalPoint[55].Cond1Cfg := 0 ;
   DigitalPoint[55].Cond2Cfg := 0 ;
   DigitalPoint[55].FlashingInputCfg := 0 ;
   
   (*DigitalPoint[56]: YA07 Node 0 Internal Defect - Smart
   ============================================================*)
   DigitalPoint[56].EnableCfg := 1 ;
   DigitalPoint[56].ActiveStateCFg := 1 ;
   DigitalPoint[56].RealInputCfg := 0 ;
   DigitalPoint[56].InputAddressCfg := 56 ;
   DigitalPoint[56].AlarmCfg := 1 ;
   DigitalPoint[56].AlarmStateCfg := 1 ;
   DigitalPoint[56].OverrideCfg := 1 ;
   DigitalPoint[56].PriorityCfg := 1 ;
   DigitalPoint[56].Cond1Cfg := 0 ;
   DigitalPoint[56].Cond2Cfg := 0 ;
   DigitalPoint[56].FlashingInputCfg := 0 ;
   
   (*DigitalPoint[57]: YA08 Node 1 Communication Failure - Clamshell
   ============================================================*)
   DigitalPoint[57].EnableCfg := 1 ;
   DigitalPoint[57].ActiveStateCFg := 1 ;
   DigitalPoint[57].RealInputCfg := 0 ;
   DigitalPoint[57].InputAddressCfg := 57 ;
   DigitalPoint[57].AlarmCfg := 1 ;
   DigitalPoint[57].AlarmStateCfg := 1 ;
   DigitalPoint[57].OverrideCfg := 1 ;
   DigitalPoint[57].PriorityCfg := 1 ;
   DigitalPoint[57].Cond1Cfg := 0 ;
   DigitalPoint[57].Cond2Cfg := 0 ;
   DigitalPoint[57].FlashingInputCfg := 0 ;
   
   (*DigitalPoint[58]: YA09 Node 1 Internal Defect - Clamshell
   ============================================================*)
   DigitalPoint[58].EnableCfg := 1 ;
   DigitalPoint[58].ActiveStateCFg := 1 ;
   DigitalPoint[58].RealInputCfg := 0 ;
   DigitalPoint[58].InputAddressCfg := 58 ;
   DigitalPoint[58].AlarmCfg := 1 ;
   DigitalPoint[58].AlarmStateCfg := 1 ;
   DigitalPoint[58].OverrideCfg := 1 ;
   DigitalPoint[58].PriorityCfg := 1 ;
   DigitalPoint[58].Cond1Cfg := 0 ;
   DigitalPoint[58].Cond2Cfg := 0 ;
   DigitalPoint[58].FlashingInputCfg := 0 ;
   
   (*DigitalPoint[59]: YA10 PLC Program Major Fault
   ============================================================*)
   DigitalPoint[59].EnableCfg := 1 ;
   DigitalPoint[59].ActiveStateCFg := 0 ;
   DigitalPoint[59].RealInputCfg := 0 ;
   DigitalPoint[59].InputAddressCfg := 59 ;
   DigitalPoint[59].AlarmCfg := 1 ;
   DigitalPoint[59].AlarmStateCfg := 1 ;
   DigitalPoint[59].OverrideCfg := 0 ;
   DigitalPoint[59].Priority := 1 ;
   DigitalPoint[59].PriorityCfg := 0 ;
   DigitalPoint[59].Cond1Cfg := 0 ;
   DigitalPoint[59].Cond2Cfg := 0 ;
   DigitalPoint[59].FlashingInputCfg := 0 ;
   
   (*DigitalPoint[60]: YA11 Database Corrupted
   ============================================================*)
   DigitalPoint[60].EnableCfg := 1 ;
   DigitalPoint[60].ActiveStateCFg := 1 ;
   DigitalPoint[60].RealInputCfg := 0 ;
   DigitalPoint[60].InputAddressCfg := 60 ;
   DigitalPoint[60].AlarmCfg := 1 ;
   DigitalPoint[60].AlarmStateCfg := 1 ;
   DigitalPoint[60].OverrideCfg := 1 ;
   DigitalPoint[60].PriorityCfg := 1 ;
   DigitalPoint[60].Cond1Cfg := 0 ;
   DigitalPoint[60].Cond2Cfg := 0 ;
   DigitalPoint[60].FlashingInputCfg := 0 ;
   
   (*DigitalPoint[61]: YA12 Unauthorized accesses
   ============================================================*)
   DigitalPoint[61].EnableCfg := 1 ;
   DigitalPoint[61].ActiveStateCFg := 1 ;
   DigitalPoint[61].RealInputCfg := 0 ;
   DigitalPoint[61].InputAddressCfg := 61 ;
   DigitalPoint[61].AlarmCfg := 1 ;
   DigitalPoint[61].AlarmStateCfg := 1 ;
   DigitalPoint[61].OverrideCfg := 1 ;
   DigitalPoint[61].PriorityCfg := 1 ;
   DigitalPoint[61].Cond1Cfg := 0 ;
   DigitalPoint[61].Cond2Cfg := 0 ;
   DigitalPoint[61].FlashingInputCfg := 0 ;
   
   (*DigitalPoint[62]: YA13 Tank Size Mismatch
   ============================================================*)
   DigitalPoint[62].EnableCfg := 1 ;
   DigitalPoint[62].ActiveStateCFg := 1 ;
   DigitalPoint[62].RealInputCfg := 0 ;
   DigitalPoint[62].InputAddressCfg := 62 ;
   DigitalPoint[62].AlarmCfg := 1 ;
   DigitalPoint[62].AlarmStateCfg := 1 ;
   DigitalPoint[62].OverrideCfg := 1 ;
   DigitalPoint[62].PriorityCfg := 1 ;
   DigitalPoint[62].Cond1Cfg := 0 ;
   DigitalPoint[62].Cond2Cfg := 0 ;
   DigitalPoint[62].FlashingInputCfg := 0 ;
   
   (*DigitalPoint[63]: YA14 SQL Server Write Failure
   ============================================================*)
   DigitalPoint[63].EnableCfg := 1 ;
   DigitalPoint[63].ActiveStateCFg := 0 ;
   DigitalPoint[63].RealInputCfg := 0 ;
   DigitalPoint[63].InputAddressCfg := 63 ;
   DigitalPoint[63].AlarmCfg := 1 ;
   DigitalPoint[63].AlarmStateCfg := 1 ;
   DigitalPoint[63].OverrideCfg := 0 ;
   DigitalPoint[63].PriorityCfg := 0 ;
   DigitalPoint[63].Priority := 0 ;
   DigitalPoint[63].Cond1Cfg := 0 ;
   DigitalPoint[63].Cond2Cfg := 0 ;
   DigitalPoint[63].FlashingInputCfg := 0 ;
   
   (*DigitalPoint[64]: UserNCr1 User Non Critical Alarm 1
   ============================================================*)
   DigitalPoint[64].EnableCfg := 1 ;
   DigitalPoint[64].ActiveStateCFg := 0 ;
   DigitalPoint[64].RealInputCfg := 0 ;
   DigitalPoint[64].InputAddressCfg := 64 ;
   DigitalPoint[64].AlarmCfg := 0 ;
   DigitalPoint[64].AlarmStateCfg := 0 ;
   DigitalPoint[64].OverrideCfg := 0 ;
   DigitalPoint[64].Override := 0 ;
   DigitalPoint[64].PriorityCfg := 0 ;
   DigitalPoint[64].Priority := 0 ;
   DigitalPoint[64].Cond1Cfg := 0 ;
   DigitalPoint[64].Cond2Cfg := 0 ;
   DigitalPoint[64].FlashingInputCfg := 0 ;
   
   (*DigitalPoint[65]: UserCr1 User Critical Alarm 1
   ============================================================*)
   DigitalPoint[65].EnableCfg := 1 ;
   DigitalPoint[65].ActiveStateCFg := 0 ;
   DigitalPoint[65].RealInputCfg := 0 ;
   DigitalPoint[65].InputAddressCfg := 65 ;
   DigitalPoint[65].AlarmCfg := 0 ;
   DigitalPoint[65].AlarmStateCfg := 0 ;
   DigitalPoint[65].OverrideCfg := 0 ;
   DigitalPoint[65].Override := 0 ;
   DigitalPoint[65].PriorityCfg := 0 ;
   DigitalPoint[65].Priority := 1 ;
   DigitalPoint[65].Cond1Cfg := 0 ;
   DigitalPoint[65].Cond2Cfg := 0 ;
   DigitalPoint[65].FlashingInputCfg := 0 ;
   
   (*DigitalPoint[66]: UserNCr2 User Non Critical Alarm 2
   ============================================================*)
   DigitalPoint[66].EnableCfg := 1 ;
   DigitalPoint[66].ActiveStateCFg := 0 ;
   DigitalPoint[66].RealInputCfg := 0 ;
   DigitalPoint[66].InputAddressCfg := 66 ;
   DigitalPoint[66].AlarmCfg := 0 ;
   DigitalPoint[66].AlarmStateCfg := 0 ;
   DigitalPoint[66].OverrideCfg := 0 ;
   DigitalPoint[66].Override := 0 ;
   DigitalPoint[66].PriorityCfg := 0 ;
   DigitalPoint[66].Priority := 0 ;
   DigitalPoint[66].Cond1Cfg := 0 ;
   DigitalPoint[66].Cond2Cfg := 0 ;
   DigitalPoint[66].FlashingInputCfg := 0 ;
   
   (*DigitalPoint[67]: UserCr2 User Critical Alarm 2
   ============================================================*)
   DigitalPoint[67].EnableCfg := 1 ;
   DigitalPoint[67].ActiveStateCFg := 0 ;
   DigitalPoint[67].RealInputCfg := 0 ;
   DigitalPoint[67].InputAddressCfg := 67 ;
   DigitalPoint[67].AlarmCfg := 0 ;
   DigitalPoint[67].AlarmStateCfg := 0 ;
   DigitalPoint[67].OverrideCfg := 0 ;
   DigitalPoint[67].Override := 0 ;
   DigitalPoint[67].PriorityCfg := 0 ;
   DigitalPoint[67].Priority := 1 ;
   DigitalPoint[67].Cond1Cfg := 0 ;
   DigitalPoint[67].Cond2Cfg := 0 ;
   DigitalPoint[67].FlashingInputCfg := 0 ;
   
   
   (*DigitalPoint[68]: ZSDF Clamshell Locking Defect
   ============================================================*)
   DigitalPoint[68].EnableCfg := 1 ;
   DigitalPoint[68].ActiveStateCFg := 1 ;
   DigitalPoint[68].RealInputCfg := 0 ;
   DigitalPoint[68].InputAddressCfg := 68 ;
   DigitalPoint[68].AlarmCfg := 1 ;
   DigitalPoint[68].AlarmStateCfg := 1 ;
   DigitalPoint[68].OverrideCfg := 1 ;
   DigitalPoint[68].PriorityCfg := 1 ;
   DigitalPoint[68].Cond1Cfg := 0 ;
   DigitalPoint[68].Cond2Cfg := 0 ;
   DigitalPoint[68].FlashingInputCfg := 0 ;
   
   (*DigitalPoint[69]: YA15 Node 3 Communication Failure - Pump
   ============================================================*)
   DigitalPoint[69].EnableCfg := 1 ;
   DigitalPoint[69].ActiveStateCFg := 1 ;
   DigitalPoint[69].RealInputCfg := 0 ;
   DigitalPoint[69].InputAddressCfg := 69 ;
   DigitalPoint[69].AlarmCfg := 1 ;
   DigitalPoint[69].AlarmStateCfg := 1 ;
   DigitalPoint[69].OverrideCfg := 1 ;
   DigitalPoint[69].PriorityCfg := 1 ;
   DigitalPoint[69].Cond1Cfg := 0 ;
   DigitalPoint[69].Cond2Cfg := 0 ;
   DigitalPoint[69].FlashingInputCfg := 0 ;
   
   (*DigitalPoint[70]: YA16 Node 3 Internal Defect - Pump
   ============================================================*)
   DigitalPoint[70].EnableCfg := 1 ;
   DigitalPoint[70].ActiveStateCFg := 1 ;
   DigitalPoint[70].RealInputCfg := 0 ;
   DigitalPoint[70].InputAddressCfg := 70 ;
   DigitalPoint[70].AlarmCfg := 1 ;
   DigitalPoint[70].AlarmStateCfg := 1 ;
   DigitalPoint[70].OverrideCfg := 1 ;
   DigitalPoint[70].PriorityCfg := 1 ;
   DigitalPoint[70].Cond1Cfg := 0 ;
   DigitalPoint[70].Cond2Cfg := 0 ;
   DigitalPoint[70].FlashingInputCfg := 0 ;
   
   (*DigitalPoint[71]: YA17 Node 4 Communication Failure - Instrum
   ============================================================*)
   DigitalPoint[71].EnableCfg := 1 ;
   DigitalPoint[71].ActiveStateCFg := 1 ;
   DigitalPoint[71].RealInputCfg := 0 ;
   DigitalPoint[71].InputAddressCfg := 71 ;
   DigitalPoint[71].AlarmCfg := 1 ;
   DigitalPoint[71].AlarmStateCfg := 1 ;
   DigitalPoint[71].OverrideCfg := 1 ;
   DigitalPoint[71].PriorityCfg := 1 ;
   DigitalPoint[71].Cond1Cfg := 0 ;
   DigitalPoint[71].Cond2Cfg := 0 ;
   DigitalPoint[71].FlashingInputCfg := 0 ;
   
   (*DigitalPoint[72]: YA18 Node 4 Internal Defect - Instrum
   ============================================================*)
   DigitalPoint[72].EnableCfg := 1 ;
   DigitalPoint[72].ActiveStateCFg := 1 ;
   DigitalPoint[72].RealInputCfg := 0 ;
   DigitalPoint[72].InputAddressCfg := 72 ;
   DigitalPoint[72].AlarmCfg := 1 ;
   DigitalPoint[72].AlarmStateCfg := 1 ;
   DigitalPoint[72].OverrideCfg := 1 ;
   DigitalPoint[72].PriorityCfg := 1 ;
   DigitalPoint[72].Cond1Cfg := 0 ;
   DigitalPoint[72].Cond2Cfg := 0 ;
   DigitalPoint[72].FlashingInputCfg := 0 ;
   
   (*DigitalPoint[73]: YA19 Node 5 Communication Failure - Tank
   ============================================================*)
   DigitalPoint[73].EnableCfg := 1 ;
   DigitalPoint[73].ActiveStateCFg := 1 ;
   DigitalPoint[73].RealInputCfg := 0 ;
   DigitalPoint[73].InputAddressCfg := 73 ;
   DigitalPoint[73].AlarmCfg := 1 ;
   DigitalPoint[73].AlarmStateCfg := 1 ;
   DigitalPoint[73].OverrideCfg := 1 ;
   DigitalPoint[73].PriorityCfg := 1 ;
   DigitalPoint[73].Cond1Cfg := 0 ;
   DigitalPoint[73].Cond2Cfg := 0 ;
   DigitalPoint[73].FlashingInputCfg := 0 ;
   
   (*DigitalPoint[74]: YA20 Node 5 Internal Defect - Tank
   ============================================================*)
   DigitalPoint[74].EnableCfg := 1 ;
   DigitalPoint[74].ActiveStateCFg := 1 ;
   DigitalPoint[74].RealInputCfg := 0 ;
   DigitalPoint[74].InputAddressCfg := 74 ;
   DigitalPoint[74].AlarmCfg := 1 ;
   DigitalPoint[74].AlarmStateCfg := 1 ;
   DigitalPoint[74].OverrideCfg := 1 ;
   DigitalPoint[74].PriorityCfg := 1 ;
   DigitalPoint[74].Cond1Cfg := 0 ;
   DigitalPoint[74].Cond2Cfg := 0 ;
   DigitalPoint[74].FlashingInputCfg := 0 ;
   
   (*DigitalPoint[75]: YA21 IND331 Communication Failure
   ============================================================*)
   DigitalPoint[75].EnableCfg := 1 ;
   DigitalPoint[75].ActiveStateCFg := 1 ;
   DigitalPoint[75].RealInputCfg := 0 ;
   DigitalPoint[75].InputAddressCfg := 75 ;
   DigitalPoint[75].AlarmCfg := 1 ;
   DigitalPoint[75].AlarmStateCfg := 1 ;
   DigitalPoint[75].OverrideCfg := 1 ;
   DigitalPoint[75].PriorityCfg := 1 ;
   DigitalPoint[75].Cond1Cfg := 0 ;
   DigitalPoint[75].Cond2Cfg := 0 ;
   DigitalPoint[75].FlashingInputCfg := 0 ;
   
   (*DigitalPoint[76]: YA22 IND131 Communication Failure
   ============================================================*)
   
   IF Options.No_Filtrate_Measurement OR Options.WI102 OR Options.FI101 OR Options.WI102_FI101 THEN
   	DigitalPoint[76].EnableCfg := 0 ;
   	DigitalPoint[76].AlarmCfg := 0 ;
   	DigitalPoint[76].Alarm := 0 ;
   ELSIF Options.WI101 OR Options.WI101_FI101 THEN
   	DigitalPoint[76].EnableCfg := 1 ;
   	DigitalPoint[76].AlarmCfg := 1 ;
   ELSE
   	DigitalPoint[76].EnableCfg := 0 ;
   	DigitalPoint[76].AlarmCfg := 0 ;
   	DigitalPoint[76].Alarm := 0 ;
   END_IF;
   
   DigitalPoint[76].ActiveStateCFg := 1 ;
   DigitalPoint[76].RealInputCfg := 0 ;
   DigitalPoint[76].InputAddressCfg := 76 ;
   DigitalPoint[76].AlarmStateCfg := 1 ;
   DigitalPoint[76].OverrideCfg := 1 ;
   DigitalPoint[76].PriorityCfg := 1 ;
   DigitalPoint[76].Cond1Cfg := 0 ;
   DigitalPoint[76].Cond2Cfg := 0 ;
   DigitalPoint[76].FlashingInputCfg := 0 ;
   
   (*DigitalPoint[77]: YA41 Operating Time Exceeded - Always non critical
   ============================================================*)
   DigitalPoint[77].EnableCfg := 1 ;
   DigitalPoint[77].ActiveStateCFg := 1 ;
   DigitalPoint[77].RealInputCfg := 0 ;
   DigitalPoint[77].InputAddressCfg := 77 ;
   DigitalPoint[77].AlarmCfg := 1 ;
   DigitalPoint[77].AlarmStateCfg := 1 ;
   DigitalPoint[77].OverrideCfg := 1 ;
   DigitalPoint[77].PriorityCfg := 0 ;
   DigitalPoint[77].Cond1Cfg := 0 ;
   DigitalPoint[77].Cond2Cfg := 0 ;
   DigitalPoint[77].FlashingInputCfg := 0 ;
   
   (*Reset Loop : Set to 0 the DigitalPoint[78 to 89].EnableCfg
   ============================================================*)
   FOR Config.IndexDP := 78 to 89 by 1 do
   	DigitalPoint[Config.IndexDP].EnableCfg := 0 ;
   	DigitalPoint[Config.IndexDP].AlarmCfg := 0 ;
   End_for ;
   
   (*DigitalPoint[90]: AI101_SIG Filtrate Conductivity Signal default
   ============================================================*)
   
   IF Options.No_Device_Connected OR Options.AI102_AI103 THEN
   	DigitalPoint[90].EnableCfg := 0 ;
   	DigitalPoint[90].AlarmCfg := 0 ;
   	DigitalPoint[90].Alarm := 0 ;
   ELSIF Options.AI101 OR Options.AI101_AI102_AI103  OR Options.AI101_AI104 OR Options.AI101_AI102_AI103_AI104 THEN
   	DigitalPoint[90].EnableCfg := 1 ;
   	DigitalPoint[90].AlarmCfg := 1 ;
   ELSE
   	DigitalPoint[90].EnableCfg := 0 ;
   	DigitalPoint[90].AlarmCfg := 0 ;
   	DigitalPoint[90].Alarm := 0 ;
   END_IF;
   
   DigitalPoint[90].ActiveStateCFg := 1 ;
   DigitalPoint[90].RealInputCfg := 0 ;
   DigitalPoint[90].InputAddressCfg := 90 ;
   DigitalPoint[90].AlarmStateCfg := 1 ;
   DigitalPoint[90].OverrideCfg := 1 ;
   DigitalPoint[90].PriorityCfg := 1 ;
   DigitalPoint[90].Cond1Cfg := 0 ;
   DigitalPoint[90].Cond2Cfg := 0 ;
   DigitalPoint[90].FlashingInputCfg := 0 ;
   
   (*DigitalPoint[91]: AI102_SIG Filtrate UV Signal default
   ============================================================*)
   
   IF Options.No_Device_Connected OR Options.AI101 OR Options.AI101_AI104 THEN
   	DigitalPoint[91].EnableCfg := 0 ;
   	DigitalPoint[91].AlarmCfg := 0 ;
   	DigitalPoint[91].Alarm := 0 ;
   ELSIF Options.AI102_AI103 OR Options.AI101_AI102_AI103 OR Options.AI101_AI102_AI103_AI104 THEN
   	DigitalPoint[91].EnableCfg := 1 ;
   	DigitalPoint[91].AlarmCfg := 1 ;
   ELSE
   	DigitalPoint[91].EnableCfg := 0 ;
   	DigitalPoint[91].AlarmCfg := 0 ;
   	DigitalPoint[91].Alarm := 0 ;
   END_IF;
   
   DigitalPoint[91].ActiveStateCFg := 1 ;
   DigitalPoint[91].RealInputCfg := 0 ;
   DigitalPoint[91].InputAddressCfg := 91 ;
   DigitalPoint[91].AlarmStateCfg := 1 ;
   DigitalPoint[91].OverrideCfg := 1 ;
   DigitalPoint[91].PriorityCfg := 1 ;
   DigitalPoint[91].Cond1Cfg := 0 ;
   DigitalPoint[91].Cond2Cfg := 0 ;
   DigitalPoint[91].FlashingInputCfg := 0 ;
   
   (*DigitalPoint[92]: AI103_SIG Filtrate UV Signal default
   ============================================================*)
   
   IF Options.No_Device_Connected OR Options.AI101 OR Options.AI101_AI104 THEN
   	DigitalPoint[92].EnableCfg := 0 ;
   	DigitalPoint[92].AlarmCfg := 0 ;
   	DigitalPoint[92].Alarm := 0 ;
   ELSIF Options.AI102_AI103 OR Options.AI101_AI102_AI103 OR Options.AI101_AI102_AI103_AI104 THEN
   	DigitalPoint[92].EnableCfg := 1 ;
   	DigitalPoint[92].AlarmCfg := 1 ;
   ELSE
   	DigitalPoint[92].EnableCfg := 0 ;
   	DigitalPoint[92].AlarmCfg := 0 ;
   	DigitalPoint[92].Alarm := 0 ;
   END_IF;
   
   DigitalPoint[92].ActiveStateCFg := 1 ;
   DigitalPoint[92].RealInputCfg := 0 ;
   DigitalPoint[92].InputAddressCfg := 92 ;
   DigitalPoint[92].AlarmStateCfg := 1 ;
   DigitalPoint[92].OverrideCfg := 1 ;
   DigitalPoint[92].PriorityCfg := 1 ;
   DigitalPoint[92].Cond1Cfg := 0 ;
   DigitalPoint[92].Cond2Cfg := 0 ;
   DigitalPoint[92].FlashingInputCfg := 0 ;
   
   (*DigitalPoint[93]: FI101_SIG Filtrate Flow flow Signal default
   ============================================================*)
   
   IF Options.No_Filtrate_Measurement OR Options.WI102 OR Options.WI101 THEN
   	DigitalPoint[93].EnableCfg := 0 ;
   	DigitalPoint[93].AlarmCfg := 0 ;
   	DigitalPoint[93].Alarm := 0 ;
   ELSIF Options.FI101 OR Options.WI101_FI101 OR Options.WI102_FI101 THEN
   	DigitalPoint[93].EnableCfg := 1 ;
   	DigitalPoint[93].AlarmCfg := 1 ;
   ELSE
   	DigitalPoint[93].EnableCfg := 0 ;
   	DigitalPoint[93].AlarmCfg := 0 ;
   	DigitalPoint[93].Alarm := 0 ;
   END_IF;
   
   DigitalPoint[93].ActiveStateCFg := 1 ;
   DigitalPoint[93].RealInputCfg := 0 ;
   DigitalPoint[93].InputAddressCfg := 93 ;
   DigitalPoint[93].AlarmStateCfg := 1 ;
   DigitalPoint[93].OverrideCfg := 1 ;
   DigitalPoint[93].PriorityCfg := 1 ;
   DigitalPoint[93].Cond1Cfg := 0 ;
   DigitalPoint[93].Cond2Cfg := 0 ;
   DigitalPoint[93].FlashingInputCfg := 0 ;
   
   (*DigitalPoint[94]: WI001_SIG Feed Bag Weight Signal default
   ============================================================*)
   DigitalPoint[94].EnableCfg := 1 ;
   DigitalPoint[94].ActiveStateCFg := 1 ;
   DigitalPoint[94].RealInputCfg := 0 ;
   DigitalPoint[94].InputAddressCfg := 94 ;
   DigitalPoint[94].AlarmCfg := 1 ;
   DigitalPoint[94].AlarmStateCfg := 1 ;
   DigitalPoint[94].OverrideCfg := 1 ;
   DigitalPoint[94].PriorityCfg := 1 ;
   DigitalPoint[94].Cond1Cfg := 0 ;
   DigitalPoint[94].Cond2Cfg := 0 ;
   DigitalPoint[94].FlashingInputCfg := 0 ;
   
   (*DigitalPoint[95]: WI101_SIG Filtrate Weight Signal default
   ============================================================*)
   
   IF Options.No_Filtrate_Measurement OR Options.WI102 OR Options.FI101 OR Options.WI102_FI101 THEN
   	DigitalPoint[95].EnableCfg := 0 ;
   	DigitalPoint[95].AlarmCfg := 0 ;
   	DigitalPoint[95].Alarm := 0 ;
   ELSIF Options.WI101 OR Options.WI101_FI101 THEN
   	DigitalPoint[95].EnableCfg := 1 ;
   	DigitalPoint[95].AlarmCfg := 1 ;
   ELSE
   	DigitalPoint[95].EnableCfg := 0 ;
   	DigitalPoint[95].AlarmCfg := 0 ;
   	DigitalPoint[95].Alarm := 0 ;
   END_IF;
   
   DigitalPoint[95].ActiveStateCFg := 1 ;
   DigitalPoint[95].RealInputCfg := 0 ;
   DigitalPoint[95].InputAddressCfg := 95 ;
   DigitalPoint[95].AlarmStateCfg := 1 ;
   DigitalPoint[95].OverrideCfg := 1 ;
   DigitalPoint[95].PriorityCfg := 1 ;
   DigitalPoint[95].Cond1Cfg := 0 ;
   DigitalPoint[95].Cond2Cfg := 0 ;
   DigitalPoint[95].FlashingInputCfg := 0 ;
   
   (*DigitalPoint[96]: WI102_SIG Customer Filtrate Weight Signal default
   ============================================================*)
   
   IF Options.No_Filtrate_Measurement OR Options.WI101 OR Options.FI101 OR Options.WI101_FI101 THEN
   	DigitalPoint[96].EnableCfg := 0 ;
   	DigitalPoint[96].AlarmCfg := 0 ;
   	DigitalPoint[96].Alarm := 0 ;
   ELSIF Options.WI102 OR Options.WI102_FI101 THEN
   	DigitalPoint[96].EnableCfg := 1 ;
   	DigitalPoint[96].AlarmCfg := 1 ;
   ELSE
   	DigitalPoint[96].EnableCfg := 0 ;
   	DigitalPoint[96].AlarmCfg := 0 ;
   	DigitalPoint[96].Alarm := 0 ;
   END_IF;
   
   DigitalPoint[96].ActiveStateCFg := 1 ;
   DigitalPoint[96].RealInputCfg := 0 ;
   DigitalPoint[96].InputAddressCfg := 96 ;
   DigitalPoint[96].AlarmStateCfg := 1 ;
   DigitalPoint[96].OverrideCfg := 1 ;
   DigitalPoint[96].PriorityCfg := 1 ;
   DigitalPoint[96].Cond1Cfg := 0 ;
   DigitalPoint[96].Cond2Cfg := 0 ;
   DigitalPoint[96].FlashingInputCfg := 0 ;
   
   (*DigitalPoint[97]: PI001_SIG Feed Pressure Signal default
   ============================================================*)
   DigitalPoint[97].EnableCfg := 1 ;
   DigitalPoint[97].ActiveStateCFg := 1 ;
   DigitalPoint[97].RealInputCfg := 0 ;
   DigitalPoint[97].InputAddressCfg := 97 ;
   DigitalPoint[97].AlarmCfg := 1 ;
   DigitalPoint[97].AlarmStateCfg := 1 ;
   DigitalPoint[97].OverrideCfg := 1 ;
   DigitalPoint[97].PriorityCfg := 1 ;
   DigitalPoint[97].Cond1Cfg := 0 ;
   DigitalPoint[97].Cond2Cfg := 0 ;
   DigitalPoint[97].FlashingInputCfg := 0 ;
   
   (*DigitalPoint[98]: PI002_SIG Retentate Pressure Signal default
   ============================================================*)
   DigitalPoint[98].EnableCfg := 1 ;
   DigitalPoint[98].ActiveStateCFg := 1 ;
   DigitalPoint[98].RealInputCfg := 0 ;
   DigitalPoint[98].InputAddressCfg := 98 ;
   DigitalPoint[98].AlarmCfg := 1 ;
   DigitalPoint[98].AlarmStateCfg := 1 ;
   DigitalPoint[98].OverrideCfg := 1 ;
   DigitalPoint[98].PriorityCfg := 1 ;
   DigitalPoint[98].Cond1Cfg := 0 ;
   DigitalPoint[98].Cond2Cfg := 0 ;
   DigitalPoint[98].FlashingInputCfg := 0 ;
   
   (*DigitalPoint[99]: PI101_SIG Filtrate Pressure Signal default
   ============================================================*)
   DigitalPoint[99].EnableCfg := 1 ;
   DigitalPoint[99].ActiveStateCFg := 1 ;
   DigitalPoint[99].RealInputCfg := 0 ;
   DigitalPoint[99].InputAddressCfg := 99 ;
   DigitalPoint[99].AlarmCfg := 1 ;
   DigitalPoint[99].AlarmStateCfg := 1 ;
   DigitalPoint[99].OverrideCfg := 1 ;
   DigitalPoint[99].PriorityCfg := 1 ;
   DigitalPoint[99].Cond1Cfg := 0 ;
   DigitalPoint[99].Cond2Cfg := 0 ;
   DigitalPoint[99].FlashingInputCfg := 0 ;
   
   (*DigitalPoint[100]: PI401_SIG Transfer Pump Pressure Signal default
   ============================================================*)
   DigitalPoint[100].EnableCfg := 1 ;
   DigitalPoint[100].ActiveStateCFg := 1 ;
   DigitalPoint[100].RealInputCfg := 0 ;
   DigitalPoint[100].InputAddressCfg := 100 ;
   DigitalPoint[100].AlarmCfg := 1 ;
   DigitalPoint[100].AlarmStateCfg := 1 ;
   DigitalPoint[100].OverrideCfg := 1 ;
   DigitalPoint[100].PriorityCfg := 1 ;
   DigitalPoint[100].Cond1Cfg := 0 ;
   DigitalPoint[100].Cond2Cfg := 0 ;
   DigitalPoint[100].FlashingInputCfg := 0 ;
   
   (*DigitalPoint[101]: TI001_SIG Feed Bag Temperature Signal default
   ============================================================*)
   DigitalPoint[101].EnableCfg := 1 ;
   DigitalPoint[101].AlarmCfg := 1 ;
   DigitalPoint[101].ActiveStateCFg := 1 ;
   DigitalPoint[101].RealInputCfg := 0 ;
   DigitalPoint[101].InputAddressCfg := 101 ;
   DigitalPoint[101].AlarmStateCfg := 1 ;
   DigitalPoint[101].OverrideCfg := 1 ;
   DigitalPoint[101].PriorityCfg := 1 ;
   DigitalPoint[101].Cond1Cfg := 0 ;
   DigitalPoint[101].Cond2Cfg := 0 ;
   DigitalPoint[101].FlashingInputCfg := 0 ;
   
   (*DigitalPoint[102]: PCV001_SIG PCV001 Position Signal default
   ============================================================*)
   DigitalPoint[102].EnableCfg := 1 ;
   DigitalPoint[102].AlarmCfg := 1 ;
   DigitalPoint[102].ActiveStateCFg := 1 ;
   DigitalPoint[102].RealInputCfg := 0 ;
   DigitalPoint[102].InputAddressCfg := 102 ;
   DigitalPoint[102].AlarmStateCfg := 1 ;
   DigitalPoint[102].OverrideCfg := 1 ;
   DigitalPoint[102].PriorityCfg := 1 ;
   DigitalPoint[102].Cond1Cfg := 0 ;
   DigitalPoint[102].Cond2Cfg := 0 ;
   DigitalPoint[102].FlashingInputCfg := 0 ;
   
   (*DigitalPoint[103]: PCV101_SIG PCV101 Position Signal default
   ============================================================*)
   DigitalPoint[103].EnableCfg := 1 ;
   DigitalPoint[103].ActiveStateCFg := 1 ;
   DigitalPoint[103].RealInputCfg := 0 ;
   DigitalPoint[103].InputAddressCfg := 103 ;
   DigitalPoint[103].AlarmCfg := 1 ;
   DigitalPoint[103].AlarmStateCfg := 1 ;
   DigitalPoint[103].OverrideCfg := 1 ;
   DigitalPoint[103].PriorityCfg := 1 ;
   DigitalPoint[103].Cond1Cfg := 0 ;
   DigitalPoint[103].Cond2Cfg := 0 ;
   DigitalPoint[103].FlashingInputCfg := 0 ;
   
   
   (*DigitalPoint[104]: MIX001_SIG Mixer Speed Signal default
   ============================================================*)
   DigitalPoint[104].EnableCfg := 1 ;
   DigitalPoint[104].ActiveStateCFg := 1 ;
   DigitalPoint[104].RealInputCfg := 0 ;
   DigitalPoint[104].InputAddressCfg := 104 ;
   DigitalPoint[104].AlarmCfg := 1 ;
   DigitalPoint[104].AlarmStateCfg := 1 ;
   DigitalPoint[104].OverrideCfg := 1 ;
   DigitalPoint[104].PriorityCfg := 1 ;
   DigitalPoint[104].Cond1Cfg := 0 ;
   DigitalPoint[104].Cond2Cfg := 0 ;
   DigitalPoint[104].FlashingInputCfg := 0 ;
   
   (*DigitalPoint[105]: AI104_SIG Filtrate pH Signal default
   ============================================================*)
   
   IF Options.No_Device_Connected OR Options.AI102_AI103 OR Options.AI101 OR Options.AI101_AI102_AI103 THEN
   	DigitalPoint[105].EnableCfg := 0 ;
   	DigitalPoint[105].AlarmCfg := 0 ;
   	DigitalPoint[105].Alarm := 0 ;
   ELSIF Options.AI101_AI104 OR Options.AI101_AI102_AI103_AI104 THEN
   	DigitalPoint[105].EnableCfg := 1 ;
   	DigitalPoint[105].AlarmCfg := 1 ;
   ELSE
   	DigitalPoint[105].EnableCfg := 0 ;
   	DigitalPoint[105].AlarmCfg := 0 ;
   	DigitalPoint[105].Alarm := 0 ;
   END_IF;
   
   DigitalPoint[105].ActiveStateCFg := 1 ;
   DigitalPoint[105].RealInputCfg := 0 ;
   DigitalPoint[105].InputAddressCfg := 105 ;
   DigitalPoint[105].AlarmStateCfg := 1 ;
   DigitalPoint[105].OverrideCfg := 1 ;
   DigitalPoint[105].PriorityCfg := 1 ;
   DigitalPoint[105].Cond1Cfg := 0 ;
   DigitalPoint[105].Cond2Cfg := 0 ;
   DigitalPoint[105].FlashingInputCfg := 0 ;
   
   
   (*DigitalPoint[106]: FI003_SIG Retentate Flow Signal default
   ============================================================*)
   IF Options.FI003 THEN
   	DigitalPoint[106].EnableCfg := 1 ;
   	DigitalPoint[106].AlarmCfg := 1 ;
   ELSE
   	DigitalPoint[106].EnableCfg := 0 ;
   	DigitalPoint[106].AlarmCfg := 0 ;
   	DigitalPoint[106].Alarm := 0 ;
   END_IF;
   DigitalPoint[106].ActiveStateCFg := 1 ;
   DigitalPoint[106].RealInputCfg := 0 ;
   DigitalPoint[106].InputAddressCfg := 106 ;
   DigitalPoint[106].AlarmStateCfg := 1 ;
   DigitalPoint[106].OverrideCfg := 1 ;
   DigitalPoint[106].PriorityCfg := 1 ;
   DigitalPoint[106].Cond1Cfg := 0 ;
   DigitalPoint[106].Cond2Cfg := 0 ;
   DigitalPoint[106].FlashingInputCfg := 0 ;
   
   
   (*Reset Loop : Set to 0 the DigitalPoint[107 to 149].EnableCfg
   ============================================================*)
   FOR Config.IndexDP := 107 to 149 by 1 do
   	DigitalPoint[Config.IndexDP].EnableCfg := 0 ;
   	DigitalPoint[Config.IndexDP].AlarmCfg := 0 ;
   End_for ;
END_ROUTINE
